(* IEC 61131-3 sources: plcfuzz/testcases/beremiz_projects/random_projects (part 4) *)

(* Additional processing to handle clocks - in CODESYS, it only starts
    with rising edge and can not be placed inside IF statement *)
IF(t0_up = TRUE) THEN
    t0_reset := TRUE;
ELSIF(t0_start = TRUE AND t0_up = FALSE) THEN
    t0_up := TRUE;  t0_reset := FALSE;
END_IF
t0(IN:=t0_reset, PT:=T0_VALUE);

END_FUNCTION_BLOCK

(* ---- IndustrialAuto2.st ---- *)
FUNCTION_BLOCK FB_G4LTL

   (* Variable definition *)
   VAR_INPUT
      x0	: BOOL;
      x1	: BOOL;
   END_VAR
   VAR_OUTPUT
      y0	: BOOL;
   END_VAR
   VAR
   (* The total number of states equals to 1 *)
      cstate6	: LINT := 0;
   END_VAR

   (* Control logic *)
CASE cstate6 OF
0:
    IF ((x0 = FALSE) AND  (x1 = TRUE)) OR ((x0 = TRUE) AND  (x1 = FALSE)) THEN
        cstate6 := 0; y0 := FALSE;
    ELSIF ((x0 = FALSE) AND  (x1 = FALSE)) OR ((x0 = TRUE) AND  (x1 = TRUE)) THEN
        cstate6 := 0; y0 := TRUE;
    END_IF;
END_CASE;

END_FUNCTION_BLOCK

(* ---- IndustrialAuto3.st ---- *)
FUNCTION_BLOCK FB_G4LTL

   (* Variable definition *)
   VAR_INPUT
      x0	: BOOL;
      x1	: BOOL;
      x2	: BOOL;
      x3	: BOOL;
   END_VAR
   VAR_OUTPUT
      y0	: BOOL;
   END_VAR
   VAR
   (* The total number of states equals to 12 *)
      cstate3	: LINT := 0;
   END_VAR

   (* Control logic *)
CASE cstate3 OF
22:
    IF ((x0 = TRUE) AND  (x1 = TRUE) AND  (x2 = TRUE) AND  (x3 = FALSE)) THEN
        cstate3 := 247; y0 := FALSE;
    ELSIF ((x0 = FALSE) AND  ( TRUE ) AND  ( TRUE ) AND  ( TRUE )) OR ((x0 = TRUE) AND  ( TRUE ) AND  (x2 = FALSE) AND  ( TRUE )) THEN
        cstate3 := 22; y0 := FALSE;
    ELSIF ((x0 = TRUE) AND  (x1 = FALSE) AND  (x2 = TRUE) AND  (x3 = FALSE)) THEN
        cstate3 := 246; y0 := TRUE;
    ELSIF ((x0 = TRUE) AND  ( TRUE ) AND  (x2 = TRUE) AND  (x3 = TRUE)) THEN
        cstate3 := 29; y0 := FALSE;
    END_IF;
0:
    IF ((x0 = FALSE) AND  (x1 = FALSE) AND  (x2 = TRUE) AND  (x3 = FALSE)) THEN
        cstate3 := 0; y0 := FALSE;
    ELSIF ((x0 = FALSE) AND  (x1 = TRUE) AND  (x2 = TRUE) AND  (x3 = FALSE)) THEN
        cstate3 := 24; y0 := FALSE;
    ELSIF ((x0 = FALSE) AND  (x1 = TRUE) AND  ( TRUE ) AND  (x3 = TRUE)) OR ((x0 = TRUE) AND  (x1 = TRUE) AND  (x2 = FALSE) AND  (x3 = TRUE)) THEN
        cstate3 := 22; y0 := FALSE;
    ELSIF ((x0 = TRUE) AND  (x1 = TRUE) AND  (x2 = TRUE) AND  (x3 = FALSE)) THEN
        cstate3 := 28; y0 := FALSE;
    ELSIF (( TRUE ) AND  (x1 = TRUE) AND  (x2 = FALSE) AND  (x3 = FALSE)) THEN
        cstate3 := 20; y0 := FALSE;
    ELSIF ((x0 = TRUE) AND  (x1 = FALSE) AND  (x2 = TRUE) AND  (x3 = FALSE)) THEN
        cstate3 := 27; y0 := TRUE;
    ELSIF ((x0 = TRUE) AND  (x1 = TRUE) AND  (x2 = TRUE) AND  (x3 = TRUE)) THEN
        cstate3 := 29; y0 := FALSE;
    ELSIF (( TRUE ) AND  (x1 = FALSE) AND  (x2 = FALSE) AND  ( TRUE )) OR (( TRUE ) AND  (x1 = FALSE) AND  (x2 = TRUE) AND  (x3 = TRUE)) THEN
        cstate3 := 18; y0 := FALSE;
    END_IF;
243:
    IF ((x0 = FALSE) AND  (x1 = FALSE) AND  (x2 = TRUE) AND  (x3 = TRUE)) OR ((x0 = TRUE) AND  ( TRUE ) AND  (x2 = TRUE) AND  (x3 = TRUE)) THEN
        cstate3 := 29; y0 := FALSE;
    ELSIF (( TRUE ) AND  ( TRUE ) AND  (x2 = FALSE) AND  (x3 = FALSE)) THEN
        cstate3 := 20; y0 := FALSE;
    ELSIF ((x0 = FALSE) AND  (x1 = FALSE) AND  (x2 = FALSE) AND  (x3 = TRUE)) OR ((x0 = FALSE) AND  (x1 = TRUE) AND  ( TRUE ) AND  (x3 = TRUE)) OR ((x0 = TRUE) AND  ( TRUE ) AND  (x2 = FALSE) AND  (x3 = TRUE)) THEN
        cstate3 := 22; y0 := FALSE;
    ELSIF ((x0 = FALSE) AND  (x1 = TRUE) AND  (x2 = TRUE) AND  (x3 = FALSE)) THEN
        cstate3 := 24; y0 := FALSE;
    ELSIF ((x0 = TRUE) AND  (x1 = TRUE) AND  (x2 = TRUE) AND  (x3 = FALSE)) THEN
        cstate3 := 28; y0 := FALSE;
    ELSIF (( TRUE ) AND  (x1 = FALSE) AND  (x2 = TRUE) AND  (x3 = FALSE)) THEN
        cstate3 := 243; y0 := TRUE;
    END_IF;
24:
    IF ((x0 = TRUE) AND  ( TRUE ) AND  (x2 = TRUE) AND  (x3 = TRUE)) THEN
        cstate3 := 29; y0 := FALSE;
    ELSIF (( TRUE ) AND  ( TRUE ) AND  (x2 = FALSE) AND  (x3 = FALSE)) THEN
        cstate3 := 20; y0 := FALSE;
    ELSIF ((x0 = FALSE) AND  ( TRUE ) AND  ( TRUE ) AND  (x3 = TRUE)) OR ((x0 = TRUE) AND  ( TRUE ) AND  (x2 = FALSE) AND  (x3 = TRUE)) THEN
        cstate3 := 22; y0 := FALSE;
    ELSIF ((x0 = TRUE) AND  (x1 = TRUE) AND  (x2 = TRUE) AND  (x3 = FALSE)) THEN
        cstate3 := 28; y0 := FALSE;
    ELSIF ((x0 = TRUE) AND  (x1 = FALSE) AND  (x2 = TRUE) AND  (x3 = FALSE)) THEN
        cstate3 := 243; y0 := TRUE;
    ELSIF ((x0 = FALSE) AND  ( TRUE ) AND  (x2 = TRUE) AND  (x3 = FALSE)) THEN
        cstate3 := 24; y0 := FALSE;
    END_IF;
246:
    IF ((x0 = FALSE) AND  (x1 = FALSE) AND  (x2 = FALSE) AND  ( TRUE )) OR ((x0 = FALSE) AND  (x1 = TRUE) AND  (x2 = FALSE) AND  ( TRUE )) OR ((x0 = FALSE) AND  (x1 = TRUE) AND  (x2 = TRUE) AND  (x3 = TRUE)) OR ((x0 = TRUE) AND  ( TRUE ) AND  (x2 = FALSE) AND  ( TRUE )) THEN
        cstate3 := 22; y0 := FALSE;
    ELSIF (( TRUE ) AND  (x1 = FALSE) AND  (x2 = TRUE) AND  (x3 = FALSE)) THEN
        cstate3 := 246; y0 := TRUE;
    ELSIF ((x0 = FALSE) AND  (x1 = FALSE) AND  (x2 = TRUE) AND  (x3 = TRUE)) OR ((x0 = TRUE) AND  ( TRUE ) AND  (x2 = TRUE) AND  (x3 = TRUE)) THEN
        cstate3 := 29; y0 := FALSE;
    ELSIF ((x0 = FALSE) AND  (x1 = TRUE) AND  (x2 = TRUE) AND  (x3 = FALSE)) THEN
        cstate3 := 786; y0 := FALSE;
    ELSIF ((x0 = TRUE) AND  (x1 = TRUE) AND  (x2 = TRUE) AND  (x3 = FALSE)) THEN
        cstate3 := 247; y0 := FALSE;
    END_IF;
27:
    IF ((x0 = FALSE) AND  (x1 = TRUE) AND  (x2 = TRUE) AND  (x3 = FALSE)) THEN
        cstate3 := 24; y0 := FALSE;
    ELSIF (( TRUE ) AND  (x1 = TRUE) AND  (x2 = FALSE) AND  (x3 = FALSE)) THEN
        cstate3 := 20; y0 := FALSE;
    ELSIF ((x0 = FALSE) AND  (x1 = TRUE) AND  ( TRUE ) AND  (x3 = TRUE)) OR ((x0 = TRUE) AND  (x1 = TRUE) AND  (x2 = FALSE) AND  (x3 = TRUE)) THEN
        cstate3 := 22; y0 := FALSE;
    ELSIF ((x0 = TRUE) AND  (x1 = TRUE) AND  (x2 = TRUE) AND  (x3 = FALSE)) THEN
        cstate3 := 28; y0 := FALSE;
    ELSIF (( TRUE ) AND  (x1 = FALSE) AND  (x2 = TRUE) AND  (x3 = FALSE)) THEN
        cstate3 := 27; y0 := TRUE;
    ELSIF ((x0 = TRUE) AND  (x1 = TRUE) AND  (x2 = TRUE) AND  (x3 = TRUE)) THEN
        cstate3 := 29; y0 := FALSE;
    ELSIF (( TRUE ) AND  (x1 = FALSE) AND  (x2 = FALSE) AND  ( TRUE )) OR (( TRUE ) AND  (x1 = FALSE) AND  (x2 = TRUE) AND  (x3 = TRUE)) THEN
        cstate3 := 18; y0 := FALSE;
    END_IF;
247:
    IF ((x0 = FALSE) AND  (x1 = TRUE) AND  (x2 = TRUE) AND  (x3 = FALSE)) THEN
        cstate3 := 786; y0 := FALSE;
    ELSIF ((x0 = FALSE) AND  (x1 = FALSE) AND  (x2 = TRUE) AND  (x3 = FALSE)) OR ((x0 = TRUE) AND  (x1 = TRUE) AND  (x2 = TRUE) AND  (x3 = FALSE)) THEN
        cstate3 := 247; y0 := FALSE;
    ELSIF ((x0 = FALSE) AND  (x1 = FALSE) AND  (x2 = FALSE) AND  ( TRUE )) OR ((x0 = FALSE) AND  (x1 = TRUE) AND  (x2 = FALSE) AND  ( TRUE )) OR ((x0 = FALSE) AND  (x1 = TRUE) AND  (x2 = TRUE) AND  (x3 = TRUE)) OR ((x0 = TRUE) AND  ( TRUE ) AND  (x2 = FALSE) AND  ( TRUE )) THEN
        cstate3 := 22; y0 := FALSE;
    ELSIF ((x0 = TRUE) AND  (x1 = FALSE) AND  (x2 = TRUE) AND  (x3 = FALSE)) THEN
        cstate3 := 246; y0 := TRUE;
    ELSIF ((x0 = FALSE) AND  (x1 = FALSE) AND  (x2 = TRUE) AND  (x3 = TRUE)) OR ((x0 = TRUE) AND  ( TRUE ) AND  (x2 = TRUE) AND  (x3 = TRUE)) THEN
        cstate3 := 29; y0 := FALSE;
    END_IF;
786:
    IF ((x0 = TRUE) AND  (x1 = TRUE) AND  (x2 = TRUE) AND  (x3 = FALSE)) THEN
        cstate3 := 247; y0 := FALSE;
    ELSIF ((x0 = FALSE) AND  ( TRUE ) AND  (x2 = FALSE) AND  ( TRUE )) OR ((x0 = FALSE) AND  ( TRUE ) AND  (x2 = TRUE) AND  (x3 = TRUE)) OR ((x0 = TRUE) AND  ( TRUE ) AND  (x2 = FALSE) AND  ( TRUE )) THEN
        cstate3 := 22; y0 := FALSE;
    ELSIF ((x0 = FALSE) AND  ( TRUE ) AND  (x2 = TRUE) AND  (x3 = FALSE)) THEN
        cstate3 := 786; y0 := FALSE;
    ELSIF ((x0 = TRUE) AND  (x1 = FALSE) AND  (x2 = TRUE) AND  (x3 = FALSE)) THEN
        cstate3 := 246; y0 := TRUE;
    ELSIF ((x0 = TRUE) AND  ( TRUE ) AND  (x2 = TRUE) AND  (x3 = TRUE)) THEN
        cstate3 := 29; y0 := FALSE;
    END_IF;
28:
    IF ((x0 = FALSE) AND  (x1 = FALSE) AND  (x2 = TRUE) AND  (x3 = FALSE)) OR ((x0 = TRUE) AND  (x1 = TRUE) AND  (x2 = TRUE) AND  (x3 = FALSE)) THEN
        cstate3 := 28; y0 := FALSE;
    ELSIF (( TRUE ) AND  ( TRUE ) AND  (x2 = FALSE) AND  (x3 = FALSE)) THEN
        cstate3 := 20; y0 := FALSE;
    ELSIF ((x0 = FALSE) AND  (x1 = FALSE) AND  (x2 = FALSE) AND  (x3 = TRUE)) OR ((x0 = FALSE) AND  (x1 = TRUE) AND  ( TRUE ) AND  (x3 = TRUE)) OR ((x0 = TRUE) AND  ( TRUE ) AND  (x2 = FALSE) AND  (x3 = TRUE)) THEN
        cstate3 := 22; y0 := FALSE;
    ELSIF ((x0 = FALSE) AND  (x1 = TRUE) AND  (x2 = TRUE) AND  (x3 = FALSE)) THEN
        cstate3 := 24; y0 := FALSE;
    ELSIF ((x0 = TRUE) AND  (x1 = FALSE) AND  (x2 = TRUE) AND  (x3 = FALSE)) THEN
        cstate3 := 243; y0 := TRUE;
    ELSIF ((x0 = FALSE) AND  (x1 = FALSE) AND  (x2 = TRUE) AND  (x3 = TRUE)) OR ((x0 = TRUE) AND  ( TRUE ) AND  (x2 = TRUE) AND  (x3 = TRUE)) THEN
        cstate3 := 29; y0 := FALSE;
    END_IF;
29:
    IF ((x0 = TRUE) AND  (x1 = TRUE) AND  (x2 = TRUE) AND  (x3 = FALSE)) THEN
        cstate3 := 247; y0 := FALSE;
    ELSIF ((x0 = FALSE) AND  (x1 = FALSE) AND  (x2 = TRUE) AND  ( TRUE )) OR ((x0 = TRUE) AND  ( TRUE ) AND  (x2 = TRUE) AND  (x3 = TRUE)) THEN
        cstate3 := 29; y0 := FALSE;
    ELSIF ((x0 = TRUE) AND  (x1 = FALSE) AND  (x2 = TRUE) AND  (x3 = FALSE)) THEN
        cstate3 := 246; y0 := TRUE;
    ELSIF ((x0 = FALSE) AND  (x1 = FALSE) AND  (x2 = FALSE) AND  ( TRUE )) OR ((x0 = FALSE) AND  (x1 = TRUE) AND  ( TRUE ) AND  ( TRUE )) OR ((x0 = TRUE) AND  ( TRUE ) AND  (x2 = FALSE) AND  ( TRUE )) THEN
        cstate3 := 22; y0 := FALSE;
    END_IF;
18:
    IF ((x0 = TRUE) AND  (x1 = TRUE) AND  (x2 = TRUE) AND  (x3 = TRUE)) THEN
        cstate3 := 29; y0 := FALSE;
    ELSIF ((x0 = TRUE) AND  (x1 = FALSE) AND  (x2 = TRUE) AND  (x3 = FALSE)) THEN
        cstate3 := 27; y0 := TRUE;
    ELSIF ((x0 = FALSE) AND  (x1 = FALSE) AND  ( TRUE ) AND  ( TRUE )) OR ((x0 = TRUE) AND  (x1 = FALSE) AND  (x2 = FALSE) AND  ( TRUE )) OR ((x0 = TRUE) AND  (x1 = FALSE) AND  (x2 = TRUE) AND  (x3 = TRUE)) THEN
        cstate3 := 18; y0 := FALSE;
    ELSIF ((x0 = FALSE) AND  (x1 = TRUE) AND  ( TRUE ) AND  (x3 = FALSE)) OR ((x0 = TRUE) AND  (x1 = TRUE) AND  (x2 = FALSE) AND  (x3 = FALSE)) THEN
        cstate3 := 20; y0 := FALSE;
    ELSIF ((x0 = FALSE) AND  (x1 = TRUE) AND  ( TRUE ) AND  (x3 = TRUE)) OR ((x0 = TRUE) AND  (x1 = TRUE) AND  (x2 = FALSE) AND  (x3 = TRUE)) THEN
        cstate3 := 22; y0 := FALSE;
    ELSIF ((x0 = TRUE) AND  (x1 = TRUE) AND  (x2 = TRUE) AND  (x3 = FALSE)) THEN
        cstate3 := 28; y0 := FALSE;
    END_IF;
20:
    IF ((x0 = TRUE) AND  ( TRUE ) AND  (x2 = TRUE) AND  (x3 = TRUE)) THEN
        cstate3 := 29; y0 := FALSE;
    ELSIF ((x0 = FALSE) AND  ( TRUE ) AND  ( TRUE ) AND  (x3 = TRUE)) OR ((x0 = TRUE) AND  ( TRUE ) AND  (x2 = FALSE) AND  (x3 = TRUE)) THEN
        cstate3 := 22; y0 := FALSE;
    ELSIF ((x0 = FALSE) AND  ( TRUE ) AND  ( TRUE ) AND  (x3 = FALSE)) OR ((x0 = TRUE) AND  ( TRUE ) AND  (x2 = FALSE) AND  (x3 = FALSE)) THEN
        cstate3 := 20; y0 := FALSE;
    ELSIF ((x0 = TRUE) AND  (x1 = TRUE) AND  (x2 = TRUE) AND  (x3 = FALSE)) THEN
        cstate3 := 28; y0 := FALSE;
    ELSIF ((x0 = TRUE) AND  (x1 = FALSE) AND  (x2 = TRUE) AND  (x3 = FALSE)) THEN
        cstate3 := 243; y0 := TRUE;
    END_IF;
END_CASE;

END_FUNCTION_BLOCK

(* ---- IndustrialAuto4.st ---- *)
FUNCTION_BLOCK FB_G4LTL

   (* Variable definition *)
   VAR_INPUT
      x0	: BOOL;
      x1	: BOOL;
      x2	: BOOL;
      x3	: BOOL;
   END_VAR
   VAR_OUTPUT
      y0	: BOOL;
      y1	: BOOL;
   END_VAR
   VAR
   (* The total number of states equals to 2 *)
      cstate21	: LINT := 0;
   END_VAR

   (* Control logic *)
CASE cstate21 OF
0:
    IF ((x0 = FALSE) AND  (x1 = FALSE) AND  (x2 = FALSE) AND  (x3 = TRUE)) THEN
        cstate21 := 0; y0 := FALSE; y1 := FALSE;
    ELSIF ((x0 = FALSE) AND  (x1 = TRUE) AND  ( TRUE ) AND  (x3 = TRUE)) OR ((x0 = TRUE) AND  (x1 = FALSE) AND  (x2 = TRUE) AND  ( TRUE )) OR ((x0 = TRUE) AND  (x1 = TRUE) AND  (x2 = FALSE) AND  (x3 = TRUE)) OR ((x0 = TRUE) AND  (x1 = TRUE) AND  (x2 = TRUE) AND  ( TRUE )) THEN
        cstate21 := 1; y0 := FALSE; y1 := FALSE;
    ELSIF ((x0 = FALSE) AND  (x1 = FALSE) AND  (x2 = FALSE) AND  (x3 = FALSE)) OR ((x0 = FALSE) AND  (x1 = FALSE) AND  (x2 = TRUE) AND  ( TRUE )) OR ((x0 = FALSE) AND  (x1 = TRUE) AND  ( TRUE ) AND  (x3 = FALSE)) THEN
        cstate21 := 0; y0 := FALSE; y1 := FALSE;
    ELSIF ((x0 = TRUE) AND  (x1 = TRUE) AND  (x2 = FALSE) AND  (x3 = FALSE)) THEN
        cstate21 := 0; y0 := TRUE; y1 := TRUE;
    ELSIF ((x0 = TRUE) AND  (x1 = FALSE) AND  (x2 = FALSE) AND  (x3 = TRUE)) THEN
        cstate21 := 0; y0 := TRUE; y1 := FALSE;
    ELSIF ((x0 = TRUE) AND  (x1 = FALSE) AND  (x2 = FALSE) AND  (x3 = FALSE)) THEN
        cstate21 := 0; y0 := TRUE; y1 := FALSE;
    END_IF;
1:
    IF ((x0 = TRUE) AND  (x1 = FALSE) AND  (x2 = FALSE) AND  ( TRUE )) OR ((x0 = TRUE) AND  (x1 = TRUE) AND  (x2 = FALSE) AND  (x3 = FALSE)) THEN
        cstate21 := 1; y0 := FALSE; y1 := FALSE;
    ELSIF ((x0 = FALSE) AND  (x1 = FALSE) AND  (x2 = FALSE) AND  (x3 = FALSE)) OR ((x0 = FALSE) AND  (x1 = FALSE) AND  (x2 = TRUE) AND  ( TRUE )) OR ((x0 = FALSE) AND  (x1 = TRUE) AND  ( TRUE ) AND  (x3 = FALSE)) THEN
        cstate21 := 1; y0 := FALSE; y1 := FALSE;
    ELSIF ((x0 = FALSE) AND  (x1 = TRUE) AND  ( TRUE ) AND  (x3 = TRUE)) OR ((x0 = TRUE) AND  (x1 = FALSE) AND  (x2 = TRUE) AND  ( TRUE )) OR ((x0 = TRUE) AND  (x1 = TRUE) AND  (x2 = FALSE) AND  (x3 = TRUE)) OR ((x0 = TRUE) AND  (x1 = TRUE) AND  (x2 = TRUE) AND  ( TRUE )) THEN
        cstate21 := 1; y0 := FALSE; y1 := FALSE;
    ELSIF ((x0 = FALSE) AND  (x1 = FALSE) AND  (x2 = FALSE) AND  (x3 = TRUE)) THEN
        cstate21 := 1; y0 := FALSE; y1 := FALSE;
    END_IF;
END_CASE;

END_FUNCTION_BLOCK

(* ---- IndustrialAuto5.st ---- *)
FUNCTION_BLOCK FB_G4LTL

   (* Variable definition *)
   VAR_INPUT
      x0	: BOOL;
      x1	: BOOL;
      c1_geq500	: BOOL;
   END_VAR
   VAR_OUTPUT
      y0	: BOOL;
      c1_add1	: BOOL;
      c1_reset	: BOOL;
   END_VAR
   VAR
   (* The total number of states equals to 4 *)
      cstate18	: LINT := 0;
   END_VAR

   (* Control logic *)
CASE cstate18 OF
0:
    IF ((x0 = FALSE) AND  (x1 = TRUE) AND  (c1_geq500 = TRUE)) THEN
        cstate18 := 3; y0 := TRUE; c1_add1 := FALSE; c1_reset := TRUE;
    ELSIF ((x0 = FALSE) AND  (x1 = FALSE) AND  (c1_geq500 = TRUE)) THEN
        cstate18 := 3; y0 := TRUE; c1_add1 := FALSE; c1_reset := FALSE;
    ELSIF ((x0 = FALSE) AND  (x1 = TRUE) AND  (c1_geq500 = FALSE)) THEN
        cstate18 := 3; y0 := FALSE; c1_add1 := FALSE; c1_reset := TRUE;
    ELSIF ((x0 = FALSE) AND  (x1 = FALSE) AND  (c1_geq500 = FALSE)) THEN
        cstate18 := 3; y0 := FALSE; c1_add1 := FALSE; c1_reset := FALSE;
    ELSIF ((x0 = TRUE) AND  (x1 = TRUE) AND  ( TRUE )) THEN
        cstate18 := 1; y0 := FALSE; c1_add1 := FALSE; c1_reset := FALSE;
    ELSIF ((x0 = TRUE) AND  (x1 = FALSE) AND  (c1_geq500 = TRUE)) THEN
        cstate18 := 2; y0 := TRUE; c1_add1 := TRUE; c1_reset := FALSE;
    ELSIF ((x0 = TRUE) AND  (x1 = FALSE) AND  (c1_geq500 = FALSE)) THEN
        cstate18 := 2; y0 := FALSE; c1_add1 := TRUE; c1_reset := FALSE;
    END_IF;
1:
    IF ((x0 = TRUE) AND  (x1 = TRUE) AND  ( TRUE )) THEN
        cstate18 := 1; y0 := FALSE; c1_add1 := FALSE; c1_reset := FALSE;
    ELSIF ((x0 = FALSE) AND  ( TRUE ) AND  (c1_geq500 = FALSE)) OR ((x0 = TRUE) AND  (x1 = FALSE) AND  (c1_geq500 = FALSE)) THEN
        cstate18 := 1; y0 := FALSE; c1_add1 := FALSE; c1_reset := FALSE;
    ELSIF ((x0 = FALSE) AND  ( TRUE ) AND  (c1_geq500 = TRUE)) OR ((x0 = TRUE) AND  (x1 = FALSE) AND  (c1_geq500 = TRUE)) THEN
        cstate18 := 1; y0 := FALSE; c1_add1 := FALSE; c1_reset := FALSE;
    END_IF;
2:
    IF ((x0 = TRUE) AND  (x1 = TRUE) AND  ( TRUE )) THEN
        cstate18 := 1; y0 := FALSE; c1_add1 := FALSE; c1_reset := FALSE;
    ELSIF ((x0 = FALSE) AND  (x1 = FALSE) AND  (c1_geq500 = TRUE)) THEN
        cstate18 := 3; y0 := TRUE; c1_add1 := FALSE; c1_reset := FALSE;
    ELSIF ((x0 = FALSE) AND  (x1 = TRUE) AND  (c1_geq500 = FALSE)) THEN
        cstate18 := 3; y0 := FALSE; c1_add1 := FALSE; c1_reset := TRUE;
    ELSIF ((x0 = FALSE) AND  (x1 = TRUE) AND  (c1_geq500 = TRUE)) THEN
        cstate18 := 3; y0 := TRUE; c1_add1 := FALSE; c1_reset := TRUE;
    ELSIF ((x0 = FALSE) AND  (x1 = FALSE) AND  (c1_geq500 = FALSE)) THEN
        cstate18 := 3; y0 := FALSE; c1_add1 := FALSE; c1_reset := FALSE;
    ELSIF ((x0 = TRUE) AND  (x1 = FALSE) AND  (c1_geq500 = FALSE)) THEN
        cstate18 := 2; y0 := FALSE; c1_add1 := FALSE; c1_reset := FALSE;
    ELSIF ((x0 = TRUE) AND  (x1 = FALSE) AND  (c1_geq500 = TRUE)) THEN
        cstate18 := 2; y0 := TRUE; c1_add1 := FALSE; c1_reset := FALSE;
    END_IF;
3:
    IF ((x0 = FALSE) AND  (x1 = FALSE) AND  (c1_geq500 = FALSE)) THEN
        cstate18 := 3; y0 := FALSE; c1_add1 := FALSE; c1_reset := FALSE;
    ELSIF ((x0 = FALSE) AND  (x1 = FALSE) AND  (c1_geq500 = TRUE)) THEN
        cstate18 := 3; y0 := TRUE; c1_add1 := FALSE; c1_reset := FALSE;
    ELSIF ((x0 = FALSE) AND  (x1 = TRUE) AND  (c1_geq500 = FALSE)) THEN
        cstate18 := 3; y0 := FALSE; c1_add1 := FALSE; c1_reset := TRUE;
    ELSIF ((x0 = FALSE) AND  (x1 = TRUE) AND  (c1_geq500 = TRUE)) THEN
        cstate18 := 3; y0 := TRUE; c1_add1 := FALSE; c1_reset := TRUE;
    ELSIF ((x0 = TRUE) AND  (x1 = TRUE) AND  ( TRUE )) THEN
        cstate18 := 1; y0 := FALSE; c1_add1 := FALSE; c1_reset := FALSE;
    ELSIF ((x0 = TRUE) AND  (x1 = FALSE) AND  (c1_geq500 = FALSE)) THEN
        cstate18 := 2; y0 := FALSE; c1_add1 := TRUE; c1_reset := FALSE;
    ELSIF ((x0 = TRUE) AND  (x1 = FALSE) AND  (c1_geq500 = TRUE)) THEN
        cstate18 := 2; y0 := TRUE; c1_add1 := TRUE; c1_reset := FALSE;
    END_IF;
END_CASE;

END_FUNCTION_BLOCK

(* ---- IndustrialAuto6.st ---- *)
FUNCTION_BLOCK FB_G4LTL

   (* Variable definition *)
   VAR_INPUT
      x1	: BOOL;
   END_VAR
   VAR_OUTPUT
      y1	: BOOL;
   END_VAR
   VAR
   (* The total number of states equals to 7 *)
      cstate12	: LINT := 0;
      t	: TON;
      t_reset	: BOOL := FALSE;
      t_up	: BOOL := FALSE;
      t_start	: BOOL := FALSE;
   END_VAR

   (* Constant definition (depending on compiler, one might need to move to normal variables) *)

   (* Each time constant has a difference of 1 period (cycle-time); please substract it when needed  *)
   VAR CONST
      T_VALUE	: TIME := TIME#5s;
   END_VAR

   (* Control logic *)
CASE cstate12 OF
0:
    IF ((x1 = FALSE) AND  (t.Q = FALSE)) THEN
        cstate12 := 1; y1 := FALSE; t_start := FALSE;
    ELSIF ((x1 = TRUE) AND  ( TRUE )) THEN
        cstate12 := 3; y1 := TRUE; t_start := FALSE;
    ELSIF ((x1 = FALSE) AND  (t.Q = TRUE)) THEN
        cstate12 := 5; y1 := FALSE; t_start := FALSE;
    END_IF;
1:
    IF ((x1 = FALSE) AND  (t.Q = FALSE)) THEN
        cstate12 := 1; y1 := FALSE; t_start := FALSE;
    ELSIF ((x1 = FALSE) AND  (t.Q = TRUE)) THEN
        cstate12 := 5; y1 := FALSE; t_start := FALSE;
    ELSIF ((x1 = TRUE) AND  ( TRUE )) THEN
        cstate12 := 3; y1 := TRUE; t_start := FALSE;
    END_IF;
2:
    IF ((x1 = TRUE) AND  (t.Q = FALSE)) THEN
        cstate12 := 2; y1 := TRUE; t_start := FALSE;
    ELSIF ((x1 = TRUE) AND  (t.Q = TRUE)) THEN
        cstate12 := 3; y1 := TRUE; t_start := FALSE;
    ELSIF ((x1 = FALSE) AND  (t.Q = FALSE)) THEN
        cstate12 := 4; y1 := TRUE; t_start := TRUE; t_up := FALSE;
    ELSIF ((x1 = FALSE) AND  (t.Q = TRUE)) THEN
        cstate12 := 6; y1 := TRUE; t_start := TRUE; t_up := FALSE;
    END_IF;
3:
    IF ((x1 = FALSE) AND  (t.Q = TRUE)) THEN
        cstate12 := 6; y1 := TRUE; t_start := TRUE; t_up := FALSE;
    ELSIF ((x1 = FALSE) AND  (t.Q = FALSE)) THEN
        cstate12 := 4; y1 := TRUE; t_start := TRUE; t_up := FALSE;
    ELSIF ((x1 = TRUE) AND  ( TRUE )) THEN
        cstate12 := 3; y1 := TRUE; t_start := FALSE;
    END_IF;
4:
    IF ((x1 = FALSE) AND  (t.Q = TRUE)) THEN
        cstate12 := 5; y1 := FALSE; t_start := FALSE;
    ELSIF ((x1 = FALSE) AND  (t.Q = FALSE)) THEN
        cstate12 := 4; y1 := TRUE; t_start := FALSE;
    ELSIF ((x1 = TRUE) AND  (t.Q = FALSE)) THEN
        cstate12 := 2; y1 := TRUE; t_start := FALSE;
    ELSIF ((x1 = TRUE) AND  (t.Q = TRUE)) THEN
        cstate12 := 3; y1 := TRUE; t_start := FALSE;
    END_IF;
5:
    IF ((x1 = TRUE) AND  ( TRUE )) THEN
        cstate12 := 3; y1 := TRUE; t_start := FALSE;
    ELSIF ((x1 = FALSE) AND  (t.Q = FALSE)) THEN
        cstate12 := 1; y1 := FALSE; t_start := FALSE;
    ELSIF ((x1 = FALSE) AND  (t.Q = TRUE)) THEN
        cstate12 := 5; y1 := FALSE; t_start := FALSE;
    END_IF;
6:
    IF ((x1 = FALSE) AND  (t.Q = TRUE)) THEN
        cstate12 := 5; y1 := FALSE; t_start := FALSE;
    ELSIF ((x1 = FALSE) AND  (t.Q = FALSE)) THEN
        cstate12 := 4; y1 := TRUE; t_start := FALSE;
    ELSIF ((x1 = TRUE) AND  (t.Q = FALSE)) THEN
        cstate12 := 2; y1 := TRUE; t_start := FALSE;
    ELSIF ((x1 = TRUE) AND  (t.Q = TRUE)) THEN
        cstate12 := 3; y1 := TRUE; t_start := FALSE;
    END_IF;
END_CASE;

(* Additional processing to handle clocks - in CODESYS, it only starts
    with rising edge and can not be placed inside IF statement *)
IF(t_up = TRUE) THEN
    t_reset := TRUE;
ELSIF(t_start = TRUE AND t_up = FALSE) THEN
    t_up := TRUE;  t_reset := FALSE;
END_IF
t(IN:=t_reset, PT:=T_VALUE);

END_FUNCTION_BLOCK

(* ---- IndustrialAuto7.st ---- *)
FUNCTION_BLOCK FB_G4LTL

   (* Variable definition *)
   VAR_INPUT
      x1	: BOOL;
   END_VAR
   VAR_OUTPUT
      y1	: BOOL;
   END_VAR
   VAR
   (* The total number of states equals to 7 *)
      cstate71	: LINT := 0;
      t	: TON;
      t_reset	: BOOL := FALSE;
      t_up	: BOOL := FALSE;
      t_start	: BOOL := FALSE;
   END_VAR

   (* Constant definition (depending on compiler, one might need to move to normal variables) *)

   (* Each time constant has a difference of 1 period (cycle-time); please substract it when needed  *)
   VAR CONST
      T_VALUE	: TIME := TIME#3s;
   END_VAR

   (* Control logic *)
CASE cstate71 OF
0:
    IF ((x1 = TRUE) AND  (t.Q = FALSE)) THEN
        cstate71 := 2; y1 := FALSE; t_start := FALSE;
    ELSIF ((x1 = FALSE) AND  ( TRUE )) THEN
        cstate71 := 6; y1 := FALSE; t_start := FALSE;
    ELSIF ((x1 = TRUE) AND  (t.Q = TRUE)) THEN
        cstate71 := 2; y1 := TRUE; t_start := FALSE;
    END_IF;
1:
    IF ((x1 = TRUE) AND  (t.Q = TRUE)) THEN
        cstate71 := 2; y1 := TRUE; t_start := FALSE;
    ELSIF ((x1 = TRUE) AND  (t.Q = FALSE)) THEN
        cstate71 := 1; y1 := FALSE; t_start := FALSE;
    ELSIF ((x1 = FALSE) AND  (t.Q = TRUE)) THEN
        cstate71 := 6; y1 := FALSE; t_start := FALSE;
    ELSIF ((x1 = FALSE) AND  (t.Q = FALSE)) THEN
        cstate71 := 5; y1 := FALSE; t_start := FALSE;
    END_IF;
2:
    IF ((x1 = TRUE) AND  (t.Q = FALSE)) THEN
        cstate71 := 2; y1 := FALSE; t_start := FALSE;
    ELSIF ((x1 = TRUE) AND  (t.Q = TRUE)) THEN
        cstate71 := 2; y1 := TRUE; t_start := FALSE;
    ELSIF ((x1 = FALSE) AND  ( TRUE )) THEN
        cstate71 := 6; y1 := FALSE; t_start := FALSE;
    END_IF;
3:
    IF ((x1 = TRUE) AND  (t.Q = FALSE)) THEN
        cstate71 := 3; y1 := FALSE; t_start := FALSE;
    ELSIF ((x1 = FALSE) AND  (t.Q = FALSE)) THEN
        cstate71 := 4; y1 := FALSE; t_start := FALSE;
    ELSIF ((x1 = TRUE) AND  (t.Q = TRUE)) THEN
        cstate71 := 2; y1 := TRUE; t_start := FALSE;
    ELSIF ((x1 = FALSE) AND  (t.Q = TRUE)) THEN
        cstate71 := 6; y1 := FALSE; t_start := FALSE;
    END_IF;
4:
    IF ((x1 = FALSE) AND  (t.Q = FALSE)) THEN
        cstate71 := 4; y1 := FALSE; t_start := FALSE;
    ELSIF ((x1 = FALSE) AND  (t.Q = TRUE)) THEN
        cstate71 := 6; y1 := FALSE; t_start := FALSE;
    ELSIF ((x1 = TRUE) AND  (t.Q = FALSE)) THEN
        cstate71 := 3; y1 := FALSE; t_start := TRUE; t_up := FALSE;
    ELSIF ((x1 = TRUE) AND  (t.Q = TRUE)) THEN
        cstate71 := 1; y1 := TRUE; t_start := TRUE; t_up := FALSE;
    END_IF;
5:
    IF ((x1 = FALSE) AND  (t.Q = TRUE)) THEN
        cstate71 := 6; y1 := FALSE; t_start := FALSE;
    ELSIF ((x1 = FALSE) AND  (t.Q = FALSE)) THEN
        cstate71 := 5; y1 := FALSE; t_start := FALSE;
    ELSIF ((x1 = TRUE) AND  (t.Q = TRUE)) THEN
        cstate71 := 1; y1 := TRUE; t_start := TRUE; t_up := FALSE;
    ELSIF ((x1 = TRUE) AND  (t.Q = FALSE)) THEN
        cstate71 := 3; y1 := FALSE; t_start := TRUE; t_up := FALSE;
    END_IF;
6:
    IF ((x1 = TRUE) AND  (t.Q = TRUE)) THEN
        cstate71 := 1; y1 := TRUE; t_start := TRUE; t_up := FALSE;
    ELSIF ((x1 = TRUE) AND  (t.Q = FALSE)) THEN
        cstate71 := 3; y1 := FALSE; t_start := TRUE; t_up := FALSE;
    ELSIF ((x1 = FALSE) AND  ( TRUE )) THEN
        cstate71 := 6; y1 := FALSE; t_start := FALSE;
    END_IF;
END_CASE;

(* Additional processing to handle clocks - in CODESYS, it only starts
    with rising edge and can not be placed inside IF statement *)
IF(t_up = TRUE) THEN
    t_reset := TRUE;
ELSIF(t_start = TRUE AND t_up = FALSE) THEN
    t_up := TRUE;  t_reset := FALSE;
END_IF
t(IN:=t_reset, PT:=T_VALUE);

END_FUNCTION_BLOCK

(* ---- IndustrialAuto8.st ---- *)
FUNCTION_BLOCK FB_G4LTL

   (* Variable definition *)
   VAR_INPUT
      x1	: BOOL;
   END_VAR
   VAR_OUTPUT
      y1	: BOOL;
   END_VAR
   VAR
   (* The total number of states equals to 18 *)
      cstate78	: LINT := 0;
      t0	: TON;
      t0_reset	: BOOL := FALSE;
      t0_up	: BOOL := FALSE;
      t0_start	: BOOL := FALSE;
      t1	: TON;
      t1_reset	: BOOL := FALSE;
      t1_up	: BOOL := FALSE;
      t1_start	: BOOL := FALSE;
   END_VAR

   (* Constant definition (depending on compiler, one might need to move to normal variables) *)

   (* Each time constant has a difference of 1 period (cycle-time); please substract it when needed  *)
   VAR CONST
      T0_VALUE	: TIME := TIME#5s;
      T1_VALUE	: TIME := TIME#3s;
   END_VAR

   (* Control logic *)
CASE cstate78 OF
11:
    IF ((x1 = FALSE) AND  (t0.Q = TRUE) AND  (t1.Q = TRUE)) THEN
        cstate78 := 14; y1 := TRUE; t0_start := FALSE;t1_start := TRUE; t1_up := FALSE;
    ELSIF ((x1 = TRUE) AND  (t0.Q = TRUE) AND  ( TRUE )) THEN
        cstate78 := 10; y1 := FALSE; t0_start := FALSE;t1_start := FALSE;
    ELSIF ((x1 = TRUE) AND  (t0.Q = FALSE) AND  ( TRUE )) THEN
        cstate78 := 11; y1 := FALSE; t0_start := FALSE;t1_start := FALSE;
    ELSIF ((x1 = FALSE) AND  (t0.Q = TRUE) AND  (t1.Q = FALSE)) THEN
        cstate78 := 8; y1 := TRUE; t0_start := FALSE;t1_start := TRUE; t1_up := FALSE;
    ELSIF ((x1 = FALSE) AND  (t0.Q = FALSE) AND  ( TRUE )) THEN
        cstate78 := 1; y1 := FALSE; t0_start := FALSE;t1_start := FALSE;
    END_IF;
12:
    IF ((x1 = TRUE) AND  (t0.Q = TRUE) AND  ( TRUE )) THEN
        cstate78 := 9; y1 := FALSE; t0_start := TRUE; t0_up := FALSE;t1_start := FALSE;
    ELSIF ((x1 = FALSE) AND  ( TRUE ) AND  (t1.Q = FALSE)) THEN
        cstate78 := 16; y1 := FALSE; t0_start := FALSE;t1_start := FALSE;
    ELSIF ((x1 = TRUE) AND  (t0.Q = FALSE) AND  ( TRUE )) THEN
        cstate78 := 3; y1 := FALSE; t0_start := TRUE; t0_up := FALSE;t1_start := FALSE;
    ELSIF ((x1 = FALSE) AND  ( TRUE ) AND  (t1.Q = TRUE)) THEN
        cstate78 := 4; y1 := FALSE; t0_start := FALSE;t1_start := FALSE;
    END_IF;
13:
    IF ((x1 = TRUE) AND  (t0.Q = FALSE) AND  ( TRUE )) THEN
        cstate78 := 3; y1 := FALSE; t0_start := TRUE; t0_up := FALSE;t1_start := FALSE;
    ELSIF ((x1 = TRUE) AND  (t0.Q = TRUE) AND  ( TRUE )) THEN
        cstate78 := 9; y1 := FALSE; t0_start := TRUE; t0_up := FALSE;t1_start := FALSE;
    ELSIF ((x1 = FALSE) AND  ( TRUE ) AND  (t1.Q = TRUE)) THEN
        cstate78 := 4; y1 := FALSE; t0_start := FALSE;t1_start := FALSE;
    ELSIF ((x1 = FALSE) AND  ( TRUE ) AND  (t1.Q = FALSE)) THEN
        cstate78 := 16; y1 := FALSE; t0_start := FALSE;t1_start := FALSE;
    END_IF;
14:
    IF ((x1 = TRUE) AND  (t0.Q = FALSE) AND  (t1.Q = TRUE)) THEN
        cstate78 := 3; y1 := FALSE; t0_start := TRUE; t0_up := FALSE;t1_start := FALSE;
    ELSIF ((x1 = FALSE) AND  ( TRUE ) AND  (t1.Q = TRUE)) THEN
        cstate78 := 12; y1 := FALSE; t0_start := FALSE;t1_start := FALSE;
    ELSIF ((x1 = TRUE) AND  ( TRUE ) AND  (t1.Q = FALSE)) THEN
        cstate78 := 1; y1 := FALSE; t0_start := FALSE;t1_start := FALSE;
    ELSIF ((x1 = FALSE) AND  ( TRUE ) AND  (t1.Q = FALSE)) THEN
        cstate78 := 15; y1 := TRUE; t0_start := FALSE;t1_start := FALSE;
    ELSIF ((x1 = TRUE) AND  (t0.Q = TRUE) AND  (t1.Q = TRUE)) THEN
        cstate78 := 9; y1 := FALSE; t0_start := TRUE; t0_up := FALSE;t1_start := FALSE;
    END_IF;
15:
    IF ((x1 = TRUE) AND  (t0.Q = TRUE) AND  (t1.Q = TRUE)) THEN
        cstate78 := 9; y1 := FALSE; t0_start := TRUE; t0_up := FALSE;t1_start := FALSE;
    ELSIF ((x1 = FALSE) AND  ( TRUE ) AND  (t1.Q = TRUE)) THEN
        cstate78 := 12; y1 := FALSE; t0_start := FALSE;t1_start := FALSE;
    ELSIF ((x1 = TRUE) AND  (t0.Q = FALSE) AND  (t1.Q = TRUE)) THEN
        cstate78 := 3; y1 := FALSE; t0_start := TRUE; t0_up := FALSE;t1_start := FALSE;
    ELSIF ((x1 = TRUE) AND  ( TRUE ) AND  (t1.Q = FALSE)) THEN
        cstate78 := 1; y1 := FALSE; t0_start := FALSE;t1_start := FALSE;
    ELSIF ((x1 = FALSE) AND  ( TRUE ) AND  (t1.Q = FALSE)) THEN
        cstate78 := 15; y1 := TRUE; t0_start := FALSE;t1_start := FALSE;
    END_IF;
16:
    IF ((x1 = TRUE) AND  (t0.Q = TRUE) AND  ( TRUE )) THEN
        cstate78 := 9; y1 := FALSE; t0_start := TRUE; t0_up := FALSE;t1_start := FALSE;
    ELSIF ((x1 = FALSE) AND  ( TRUE ) AND  (t1.Q = TRUE)) THEN
        cstate78 := 4; y1 := FALSE; t0_start := FALSE;t1_start := FALSE;
    ELSIF ((x1 = FALSE) AND  ( TRUE ) AND  (t1.Q = FALSE)) THEN
        cstate78 := 16; y1 := FALSE; t0_start := FALSE;t1_start := FALSE;
    ELSIF ((x1 = TRUE) AND  (t0.Q = FALSE) AND  ( TRUE )) THEN
        cstate78 := 3; y1 := FALSE; t0_start := TRUE; t0_up := FALSE;t1_start := FALSE;
    END_IF;
17:
    IF ((x1 = FALSE) AND  ( TRUE ) AND  (t1.Q = FALSE)) THEN
        cstate78 := 8; y1 := TRUE; t0_start := FALSE;t1_start := TRUE; t1_up := FALSE;
    ELSIF ((x1 = TRUE) AND  (t0.Q = FALSE) AND  ( TRUE )) THEN
        cstate78 := 6; y1 := FALSE; t0_start := FALSE;t1_start := FALSE;
    ELSIF ((x1 = FALSE) AND  ( TRUE ) AND  (t1.Q = TRUE)) THEN
        cstate78 := 14; y1 := TRUE; t0_start := FALSE;t1_start := TRUE; t1_up := FALSE;
    ELSIF ((x1 = TRUE) AND  (t0.Q = TRUE) AND  ( TRUE )) THEN
        cstate78 := 7; y1 := FALSE; t0_start := FALSE;t1_start := FALSE;
    END_IF;
0:
    IF ((x1 = TRUE) AND  (t0.Q = FALSE) AND  ( TRUE )) THEN
        cstate78 := 17; y1 := FALSE; t0_start := FALSE;t1_start := FALSE;
    ELSIF ((x1 = FALSE) AND  ( TRUE ) AND  (t1.Q = FALSE)) THEN
        cstate78 := 2; y1 := FALSE; t0_start := FALSE;t1_start := FALSE;
    ELSIF ((x1 = FALSE) AND  ( TRUE ) AND  (t1.Q = TRUE)) THEN
        cstate78 := 13; y1 := FALSE; t0_start := FALSE;t1_start := FALSE;
    ELSIF ((x1 = TRUE) AND  (t0.Q = TRUE) AND  ( TRUE )) THEN
        cstate78 := 5; y1 := FALSE; t0_start := FALSE;t1_start := FALSE;
    END_IF;
1:
    IF (( TRUE )) THEN
        cstate78 := 1; y1 := FALSE; t0_start := FALSE;t1_start := FALSE;
    END_IF;
2:
    IF ((x1 = TRUE) AND  (t0.Q = FALSE) AND  ( TRUE )) THEN
        cstate78 := 3; y1 := FALSE; t0_start := TRUE; t0_up := FALSE;t1_start := FALSE;
    ELSIF ((x1 = FALSE) AND  ( TRUE ) AND  (t1.Q = FALSE)) THEN
        cstate78 := 16; y1 := FALSE; t0_start := FALSE;t1_start := FALSE;
    ELSIF ((x1 = TRUE) AND  (t0.Q = TRUE) AND  ( TRUE )) THEN
        cstate78 := 9; y1 := FALSE; t0_start := TRUE; t0_up := FALSE;t1_start := FALSE;
    ELSIF ((x1 = FALSE) AND  ( TRUE ) AND  (t1.Q = TRUE)) THEN
        cstate78 := 4; y1 := FALSE; t0_start := FALSE;t1_start := FALSE;
    END_IF;
3:
    IF ((x1 = FALSE) AND  (t0.Q = FALSE) AND  ( TRUE )) THEN
        cstate78 := 1; y1 := FALSE; t0_start := FALSE;t1_start := FALSE;
    ELSIF ((x1 = TRUE) AND  (t0.Q = FALSE) AND  ( TRUE )) THEN
        cstate78 := 11; y1 := FALSE; t0_start := FALSE;t1_start := FALSE;
    ELSIF ((x1 = FALSE) AND  (t0.Q = TRUE) AND  (t1.Q = TRUE)) THEN
        cstate78 := 14; y1 := TRUE; t0_start := FALSE;t1_start := TRUE; t1_up := FALSE;
    ELSIF ((x1 = FALSE) AND  (t0.Q = TRUE) AND  (t1.Q = FALSE)) THEN
        cstate78 := 8; y1 := TRUE; t0_start := FALSE;t1_start := TRUE; t1_up := FALSE;
    ELSIF ((x1 = TRUE) AND  (t0.Q = TRUE) AND  ( TRUE )) THEN
        cstate78 := 10; y1 := FALSE; t0_start := FALSE;t1_start := FALSE;
    END_IF;
4:
    IF ((x1 = FALSE) AND  ( TRUE ) AND  (t1.Q = TRUE)) THEN
        cstate78 := 4; y1 := FALSE; t0_start := FALSE;t1_start := FALSE;
    ELSIF ((x1 = TRUE) AND  (t0.Q = TRUE) AND  ( TRUE )) THEN
        cstate78 := 9; y1 := FALSE; t0_start := TRUE; t0_up := FALSE;t1_start := FALSE;
    ELSIF ((x1 = FALSE) AND  ( TRUE ) AND  (t1.Q = FALSE)) THEN
        cstate78 := 16; y1 := FALSE; t0_start := FALSE;t1_start := FALSE;
    ELSIF ((x1 = TRUE) AND  (t0.Q = FALSE) AND  ( TRUE )) THEN
        cstate78 := 3; y1 := FALSE; t0_start := TRUE; t0_up := FALSE;t1_start := FALSE;
    END_IF;
5:
    IF ((x1 = TRUE) AND  (t0.Q = FALSE) AND  ( TRUE )) THEN
        cstate78 := 6; y1 := FALSE; t0_start := FALSE;t1_start := FALSE;
    ELSIF ((x1 = FALSE) AND  ( TRUE ) AND  (t1.Q = TRUE)) THEN
        cstate78 := 14; y1 := TRUE; t0_start := FALSE;t1_start := TRUE; t1_up := FALSE;
    ELSIF ((x1 = FALSE) AND  ( TRUE ) AND  (t1.Q = FALSE)) THEN
        cstate78 := 8; y1 := TRUE; t0_start := FALSE;t1_start := TRUE; t1_up := FALSE;
    ELSIF ((x1 = TRUE) AND  (t0.Q = TRUE) AND  ( TRUE )) THEN
        cstate78 := 7; y1 := TRUE; t0_start := FALSE;t1_start := FALSE;
    END_IF;
6:
    IF ((x1 = TRUE) AND  (t0.Q = TRUE) AND  ( TRUE )) THEN
        cstate78 := 7; y1 := FALSE; t0_start := FALSE;t1_start := FALSE;
    ELSIF ((x1 = TRUE) AND  (t0.Q = FALSE) AND  ( TRUE )) THEN
        cstate78 := 6; y1 := FALSE; t0_start := FALSE;t1_start := FALSE;
    ELSIF ((x1 = FALSE) AND  ( TRUE ) AND  (t1.Q = TRUE)) THEN
        cstate78 := 14; y1 := TRUE; t0_start := FALSE;t1_start := TRUE; t1_up := FALSE;
    ELSIF ((x1 = FALSE) AND  ( TRUE ) AND  (t1.Q = FALSE)) THEN
        cstate78 := 8; y1 := TRUE; t0_start := FALSE;t1_start := TRUE; t1_up := FALSE;
    END_IF;
7:
    IF ((x1 = FALSE) AND  ( TRUE ) AND  (t1.Q = FALSE)) THEN
        cstate78 := 8; y1 := TRUE; t0_start := FALSE;t1_start := TRUE; t1_up := FALSE;
    ELSIF ((x1 = FALSE) AND  ( TRUE ) AND  (t1.Q = TRUE)) THEN
        cstate78 := 14; y1 := TRUE; t0_start := FALSE;t1_start := TRUE; t1_up := FALSE;
    ELSIF ((x1 = TRUE) AND  (t0.Q = FALSE) AND  ( TRUE )) THEN
        cstate78 := 6; y1 := FALSE; t0_start := FALSE;t1_start := FALSE;
    ELSIF ((x1 = TRUE) AND  (t0.Q = TRUE) AND  ( TRUE )) THEN
        cstate78 := 7; y1 := TRUE; t0_start := FALSE;t1_start := FALSE;
    END_IF;
8:
    IF ((x1 = TRUE) AND  (t0.Q = TRUE) AND  (t1.Q = TRUE)) THEN
        cstate78 := 9; y1 := FALSE; t0_start := TRUE; t0_up := FALSE;t1_start := FALSE;
    ELSIF ((x1 = FALSE) AND  ( TRUE ) AND  (t1.Q = TRUE)) THEN
        cstate78 := 12; y1 := FALSE; t0_start := FALSE;t1_start := FALSE;
    ELSIF ((x1 = TRUE) AND  ( TRUE ) AND  (t1.Q = FALSE)) THEN
        cstate78 := 1; y1 := FALSE; t0_start := FALSE;t1_start := FALSE;
    ELSIF ((x1 = FALSE) AND  ( TRUE ) AND  (t1.Q = FALSE)) THEN
        cstate78 := 15; y1 := TRUE; t0_start := FALSE;t1_start := FALSE;
    ELSIF ((x1 = TRUE) AND  (t0.Q = FALSE) AND  (t1.Q = TRUE)) THEN
        cstate78 := 3; y1 := FALSE; t0_start := TRUE; t0_up := FALSE;t1_start := FALSE;
    END_IF;
9:
    IF ((x1 = TRUE) AND  (t0.Q = TRUE) AND  ( TRUE )) THEN
        cstate78 := 10; y1 := TRUE; t0_start := FALSE;t1_start := FALSE;
    ELSIF ((x1 = FALSE) AND  (t0.Q = FALSE) AND  ( TRUE )) THEN
        cstate78 := 1; y1 := FALSE; t0_start := FALSE;t1_start := FALSE;
    ELSIF ((x1 = FALSE) AND  (t0.Q = TRUE) AND  (t1.Q = TRUE)) THEN
        cstate78 := 14; y1 := TRUE; t0_start := FALSE;t1_start := TRUE; t1_up := FALSE;
    ELSIF ((x1 = TRUE) AND  (t0.Q = FALSE) AND  ( TRUE )) THEN
        cstate78 := 11; y1 := FALSE; t0_start := FALSE;t1_start := FALSE;
    ELSIF ((x1 = FALSE) AND  (t0.Q = TRUE) AND  (t1.Q = FALSE)) THEN
        cstate78 := 8; y1 := TRUE; t0_start := FALSE;t1_start := TRUE; t1_up := FALSE;
    END_IF;
10:
    IF ((x1 = TRUE) AND  (t0.Q = TRUE) AND  ( TRUE )) THEN
        cstate78 := 7; y1 := TRUE; t0_start := FALSE;t1_start := FALSE;
    ELSIF ((x1 = TRUE) AND  (t0.Q = FALSE) AND  ( TRUE )) THEN
        cstate78 := 6; y1 := FALSE; t0_start := FALSE;t1_start := FALSE;
    ELSIF ((x1 = FALSE) AND  ( TRUE ) AND  (t1.Q = TRUE)) THEN
        cstate78 := 14; y1 := TRUE; t0_start := FALSE;t1_start := TRUE; t1_up := FALSE;
    ELSIF ((x1 = FALSE) AND  ( TRUE ) AND  (t1.Q = FALSE)) THEN
        cstate78 := 8; y1 := TRUE; t0_start := FALSE;t1_start := TRUE; t1_up := FALSE;
    END_IF;
END_CASE;

(* Additional processing to handle clocks - in CODESYS, it only starts
    with rising edge and can not be placed inside IF statement *)
IF(t0_up = TRUE) THEN
    t0_reset := TRUE;
ELSIF(t0_start = TRUE AND t0_up = FALSE) THEN
    t0_up := TRUE;  t0_reset := FALSE;
END_IF
t0(IN:=t0_reset, PT:=T0_VALUE);
IF(t1_up = TRUE) THEN
    t1_reset := TRUE;
ELSIF(t1_start = TRUE AND t1_up = FALSE) THEN
    t1_up := TRUE;  t1_reset := FALSE;
END_IF
t1(IN:=t1_reset, PT:=T1_VALUE);

END_FUNCTION_BLOCK

(* ---- Req1.st ---- *)
FUNCTION_BLOCK FB_G4LTL

   (* Variable definition *)
   VAR_INPUT
      req1	: BOOL;
   END_VAR
   VAR_OUTPUT
      grant1	: BOOL;
   END_VAR
   VAR
   (* The total number of states equals to 1 *)
      cstate98	: LINT := 0;
   END_VAR

   (* Control logic *)
CASE cstate98 OF
0:
    IF ((req1 = FALSE)) THEN
        cstate98 := 0; grant1 := FALSE;
    ELSIF ((req1 = TRUE)) THEN
        cstate98 := 0; grant1 := TRUE;
    END_IF;
END_CASE;

END_FUNCTION_BLOCK

(* ---- Req3.st ---- *)
FUNCTION_BLOCK FB_G4LTL

   (* Variable definition *)
   VAR_INPUT
      req	: BOOL;
      cancel	: BOOL;
      go	: BOOL;
   END_VAR
   VAR_OUTPUT
      grant	: BOOL;
   END_VAR
   VAR
   (* The total number of states equals to 22 *)
      cstate23	: LINT := 0;
   END_VAR

   (* Control logic *)
CASE cstate23 OF
11:
    IF ((req = TRUE) AND  (cancel = TRUE) AND  ( TRUE )) THEN
        cstate23 := 8; grant := FALSE;
    ELSIF ((req = TRUE) AND  (cancel = FALSE) AND  ( TRUE )) THEN
        cstate23 := 15; grant := FALSE;
    ELSIF ((req = FALSE) AND  (cancel = FALSE) AND  ( TRUE )) THEN
        cstate23 := 11; grant := FALSE;
    ELSIF ((req = FALSE) AND  (cancel = TRUE) AND  ( TRUE )) THEN
        cstate23 := 19; grant := FALSE;
    END_IF;
12:
    IF ((req = TRUE) AND  (cancel = FALSE) AND  ( TRUE )) THEN
        cstate23 := 13; grant := FALSE;
    ELSIF ((req = FALSE) AND  (cancel = FALSE) AND  ( TRUE )) THEN
        cstate23 := 6; grant := FALSE;
    ELSIF ((req = TRUE) AND  (cancel = TRUE) AND  ( TRUE )) THEN
        cstate23 := 10; grant := FALSE;
    ELSIF ((req = FALSE) AND  (cancel = TRUE) AND  ( TRUE )) THEN
        cstate23 := 20; grant := FALSE;
    END_IF;
13:
    IF ((req = FALSE) AND  (cancel = FALSE) AND  ( TRUE )) THEN
        cstate23 := 7; grant := TRUE;
    ELSIF ((req = TRUE) AND  (cancel = TRUE) AND  ( TRUE )) THEN
        cstate23 := 4; grant := TRUE;
    ELSIF ((req = TRUE) AND  (cancel = FALSE) AND  ( TRUE )) THEN
        cstate23 := 2; grant := TRUE;
    ELSIF ((req = FALSE) AND  (cancel = TRUE) AND  ( TRUE )) THEN
        cstate23 := 18; grant := TRUE;
    END_IF;
14:
    IF ((req = TRUE) AND  (cancel = TRUE) AND  ( TRUE )) THEN
        cstate23 := 4; grant := TRUE;
    ELSIF ((req = TRUE) AND  (cancel = FALSE) AND  ( TRUE )) THEN
        cstate23 := 2; grant := TRUE;
    ELSIF ((req = FALSE) AND  (cancel = TRUE) AND  ( TRUE )) THEN
        cstate23 := 18; grant := TRUE;
    ELSIF ((req = FALSE) AND  (cancel = FALSE) AND  ( TRUE )) THEN
        cstate23 := 7; grant := TRUE;
    END_IF;
15:
    IF ((req = FALSE) AND  (cancel = TRUE) AND  ( TRUE )) THEN
        cstate23 := 9; grant := FALSE;
    ELSIF ((req = TRUE) AND  (cancel = FALSE) AND  ( TRUE )) THEN
        cstate23 := 21; grant := FALSE;
    ELSIF ((req = FALSE) AND  (cancel = FALSE) AND  ( TRUE )) THEN
        cstate23 := 12; grant := FALSE;
    ELSIF ((req = TRUE) AND  (cancel = TRUE) AND  ( TRUE )) THEN
        cstate23 := 17; grant := FALSE;
    END_IF;
16:
    IF (( TRUE )) THEN
        cstate23 := 16; grant := FALSE;
    END_IF;
17:
    IF ((req = FALSE) AND  (cancel = TRUE) AND  (go = TRUE)) THEN
        cstate23 := 1; grant := FALSE;
    ELSIF ((req = TRUE) AND  (cancel = FALSE) AND  (go = TRUE)) THEN
        cstate23 := 3; grant := FALSE;
    ELSIF (( TRUE ) AND  ( TRUE ) AND  (go = FALSE)) THEN
        cstate23 := 16; grant := FALSE;
    ELSIF ((req = FALSE) AND  (cancel = FALSE) AND  (go = TRUE)) THEN
        cstate23 := 14; grant := FALSE;
    ELSIF ((req = TRUE) AND  (cancel = TRUE) AND  (go = TRUE)) THEN
        cstate23 := 5; grant := FALSE;
    END_IF;
18:
    IF ((req = FALSE) AND  (cancel = FALSE) AND  (go = TRUE)) THEN
        cstate23 := 11; grant := FALSE;
    ELSIF ((req = FALSE) AND  (cancel = TRUE) AND  (go = TRUE)) THEN
        cstate23 := 19; grant := FALSE;
    ELSIF (( TRUE ) AND  ( TRUE ) AND  (go = FALSE)) THEN
        cstate23 := 16; grant := FALSE;
    ELSIF ((req = TRUE) AND  (cancel = TRUE) AND  (go = TRUE)) THEN
        cstate23 := 8; grant := FALSE;
    ELSIF ((req = TRUE) AND  (cancel = FALSE) AND  (go = TRUE)) THEN
        cstate23 := 15; grant := FALSE;
    END_IF;
19:
    IF (( TRUE ) AND  ( TRUE ) AND  (go = FALSE)) THEN
        cstate23 := 16; grant := FALSE;
    ELSIF ((req = FALSE) AND  (cancel = TRUE) AND  (go = TRUE)) THEN
        cstate23 := 19; grant := FALSE;
    ELSIF ((req = TRUE) AND  (cancel = FALSE) AND  (go = TRUE)) THEN
        cstate23 := 15; grant := FALSE;
    ELSIF ((req = FALSE) AND  (cancel = FALSE) AND  (go = TRUE)) THEN
        cstate23 := 11; grant := FALSE;
    ELSIF ((req = TRUE) AND  (cancel = TRUE) AND  (go = TRUE)) THEN
        cstate23 := 8; grant := FALSE;
    END_IF;
0:
    IF ((req = FALSE) AND  (cancel = FALSE) AND  ( TRUE )) THEN
        cstate23 := 11; grant := FALSE;
    ELSIF ((req = FALSE) AND  (cancel = TRUE) AND  ( TRUE )) THEN
        cstate23 := 19; grant := FALSE;
    ELSIF ((req = TRUE) AND  (cancel = FALSE) AND  ( TRUE )) THEN
        cstate23 := 15; grant := FALSE;
    ELSIF ((req = TRUE) AND  (cancel = TRUE) AND  ( TRUE )) THEN
        cstate23 := 8; grant := FALSE;
    END_IF;
1:
    IF ((req = TRUE) AND  (cancel = FALSE) AND  (go = TRUE)) THEN
        cstate23 := 2; grant := TRUE;
    ELSIF ((req = FALSE) AND  (cancel = TRUE) AND  (go = TRUE)) THEN
        cstate23 := 18; grant := TRUE;
    ELSIF ((req = FALSE) AND  (cancel = FALSE) AND  (go = TRUE)) THEN
        cstate23 := 7; grant := TRUE;
    ELSIF ((req = TRUE) AND  (cancel = TRUE) AND  (go = TRUE)) THEN
        cstate23 := 4; grant := TRUE;
    ELSIF (( TRUE ) AND  ( TRUE ) AND  (go = FALSE)) THEN
        cstate23 := 16; grant := FALSE;
    END_IF;
2:
    IF ((req = FALSE) AND  (cancel = FALSE) AND  ( TRUE )) THEN
        cstate23 := 12; grant := FALSE;
    ELSIF ((req = TRUE) AND  (cancel = TRUE) AND  ( TRUE )) THEN
        cstate23 := 17; grant := FALSE;
    ELSIF ((req = FALSE) AND  (cancel = TRUE) AND  ( TRUE )) THEN
        cstate23 := 9; grant := FALSE;
    ELSIF ((req = TRUE) AND  (cancel = FALSE) AND  ( TRUE )) THEN
        cstate23 := 21; grant := FALSE;
    END_IF;
3:
    IF ((req = TRUE) AND  (cancel = TRUE) AND  ( TRUE )) THEN
        cstate23 := 4; grant := TRUE;
    ELSIF ((req = FALSE) AND  (cancel = FALSE) AND  ( TRUE )) THEN
        cstate23 := 7; grant := TRUE;
    ELSIF ((req = TRUE) AND  (cancel = FALSE) AND  ( TRUE )) THEN
        cstate23 := 2; grant := TRUE;
    ELSIF ((req = FALSE) AND  (cancel = TRUE) AND  ( TRUE )) THEN
        cstate23 := 18; grant := TRUE;
    END_IF;
4:
    IF (( TRUE ) AND  ( TRUE ) AND  (go = FALSE)) THEN
        cstate23 := 16; grant := FALSE;
    ELSIF ((req = FALSE) AND  (cancel = TRUE) AND  (go = TRUE)) THEN
        cstate23 := 9; grant := FALSE;
    ELSIF ((req = TRUE) AND  (cancel = FALSE) AND  (go = TRUE)) THEN
        cstate23 := 21; grant := FALSE;
    ELSIF ((req = FALSE) AND  (cancel = FALSE) AND  (go = TRUE)) THEN
        cstate23 := 12; grant := FALSE;
    ELSIF ((req = TRUE) AND  (cancel = TRUE) AND  (go = TRUE)) THEN
        cstate23 := 17; grant := FALSE;
    END_IF;
5:
    IF ((req = TRUE) AND  (cancel = FALSE) AND  (go = TRUE)) THEN
        cstate23 := 2; grant := TRUE;
    ELSIF ((req = FALSE) AND  (cancel = TRUE) AND  (go = TRUE)) THEN
        cstate23 := 18; grant := TRUE;
    ELSIF (( TRUE ) AND  ( TRUE ) AND  (go = FALSE)) THEN
        cstate23 := 16; grant := FALSE;
    ELSIF ((req = TRUE) AND  (cancel = TRUE) AND  (go = TRUE)) THEN
        cstate23 := 4; grant := TRUE;
    ELSIF ((req = FALSE) AND  (cancel = FALSE) AND  (go = TRUE)) THEN
        cstate23 := 7; grant := TRUE;
    END_IF;
6:
    IF ((req = FALSE) AND  (cancel = FALSE) AND  ( TRUE )) THEN
        cstate23 := 7; grant := TRUE;
    ELSIF ((req = TRUE) AND  (cancel = TRUE) AND  ( TRUE )) THEN
        cstate23 := 4; grant := TRUE;
    ELSIF ((req = TRUE) AND  (cancel = FALSE) AND  ( TRUE )) THEN
        cstate23 := 2; grant := TRUE;
    ELSIF ((req = FALSE) AND  (cancel = TRUE) AND  ( TRUE )) THEN
        cstate23 := 18; grant := TRUE;
    END_IF;
7:
    IF ((req = TRUE) AND  (cancel = TRUE) AND  ( TRUE )) THEN
        cstate23 := 8; grant := FALSE;
    ELSIF ((req = TRUE) AND  (cancel = FALSE) AND  ( TRUE )) THEN
        cstate23 := 15; grant := FALSE;
    ELSIF ((req = FALSE) AND  (cancel = FALSE) AND  ( TRUE )) THEN
        cstate23 := 11; grant := FALSE;
    ELSIF ((req = FALSE) AND  (cancel = TRUE) AND  ( TRUE )) THEN
        cstate23 := 19; grant := FALSE;
    END_IF;
8:
    IF ((req = FALSE) AND  (cancel = TRUE) AND  (go = TRUE)) THEN
        cstate23 := 9; grant := FALSE;
    ELSIF ((req = TRUE) AND  (cancel = TRUE) AND  (go = TRUE)) THEN
        cstate23 := 17; grant := FALSE;
    ELSIF ((req = FALSE) AND  (cancel = FALSE) AND  (go = TRUE)) THEN
        cstate23 := 12; grant := FALSE;
    ELSIF ((req = TRUE) AND  (cancel = FALSE) AND  (go = TRUE)) THEN
        cstate23 := 21; grant := FALSE;
    ELSIF (( TRUE ) AND  ( TRUE ) AND  (go = FALSE)) THEN
        cstate23 := 16; grant := FALSE;
    END_IF;
9:
    IF ((req = TRUE) AND  (cancel = TRUE) AND  (go = TRUE)) THEN
        cstate23 := 10; grant := FALSE;
    ELSIF ((req = FALSE) AND  (cancel = TRUE) AND  (go = TRUE)) THEN
        cstate23 := 20; grant := FALSE;
    ELSIF ((req = TRUE) AND  (cancel = FALSE) AND  (go = TRUE)) THEN
        cstate23 := 13; grant := FALSE;
    ELSIF (( TRUE ) AND  ( TRUE ) AND  (go = FALSE)) THEN
        cstate23 := 16; grant := FALSE;
    ELSIF ((req = FALSE) AND  (cancel = FALSE) AND  (go = TRUE)) THEN
        cstate23 := 6; grant := FALSE;
    END_IF;
20:
    IF ((req = TRUE) AND  (cancel = FALSE) AND  (go = TRUE)) THEN
        cstate23 := 2; grant := TRUE;
    ELSIF ((req = FALSE) AND  (cancel = TRUE) AND  (go = TRUE)) THEN
        cstate23 := 18; grant := TRUE;
    ELSIF (( TRUE ) AND  ( TRUE ) AND  (go = FALSE)) THEN
        cstate23 := 16; grant := FALSE;
    ELSIF ((req = FALSE) AND  (cancel = FALSE) AND  (go = TRUE)) THEN
        cstate23 := 7; grant := TRUE;
    ELSIF ((req = TRUE) AND  (cancel = TRUE) AND  (go = TRUE)) THEN
        cstate23 := 4; grant := TRUE;
    END_IF;
10:
    IF ((req = FALSE) AND  (cancel = FALSE) AND  (go = TRUE)) THEN
        cstate23 := 7; grant := TRUE;
    ELSIF ((req = TRUE) AND  (cancel = FALSE) AND  (go = TRUE)) THEN
        cstate23 := 2; grant := TRUE;
    ELSIF (( TRUE ) AND  ( TRUE ) AND  (go = FALSE)) THEN
        cstate23 := 16; grant := FALSE;
    ELSIF ((req = FALSE) AND  (cancel = TRUE) AND  (go = TRUE)) THEN
        cstate23 := 18; grant := TRUE;
    ELSIF ((req = TRUE) AND  (cancel = TRUE) AND  (go = TRUE)) THEN
        cstate23 := 4; grant := TRUE;
    END_IF;
21:
    IF ((req = FALSE) AND  (cancel = FALSE) AND  ( TRUE )) THEN
        cstate23 := 14; grant := FALSE;
    ELSIF ((req = TRUE) AND  (cancel = TRUE) AND  ( TRUE )) THEN
        cstate23 := 5; grant := FALSE;
    ELSIF ((req = FALSE) AND  (cancel = TRUE) AND  ( TRUE )) THEN
        cstate23 := 1; grant := FALSE;
    ELSIF ((req = TRUE) AND  (cancel = FALSE) AND  ( TRUE )) THEN
        cstate23 := 3; grant := FALSE;
    END_IF;
END_CASE;

END_FUNCTION_BLOCK

(* ---- Req4.st ---- *)
FUNCTION_BLOCK FB_G4LTL

   (* Variable definition *)
   VAR_INPUT
      req	: BOOL;
      cancel	: BOOL;
      go	: BOOL;
   END_VAR
   VAR_OUTPUT
      grant	: BOOL;
   END_VAR
   VAR
   (* The total number of states equals to 42 *)
      cstate34	: LINT := 0;
   END_VAR

   (* Control logic *)
CASE cstate34 OF
22:
    IF ((req = TRUE) AND  (cancel = FALSE) AND  ( TRUE )) THEN
        cstate34 := 26; grant := FALSE;
    ELSIF ((req = TRUE) AND  (cancel = TRUE) AND  ( TRUE )) THEN
        cstate34 := 14; grant := FALSE;
    ELSIF ((req = FALSE) AND  (cancel = FALSE) AND  ( TRUE )) THEN
        cstate34 := 7; grant := FALSE;
    ELSIF ((req = FALSE) AND  (cancel = TRUE) AND  ( TRUE )) THEN
        cstate34 := 19; grant := FALSE;
    END_IF;
23:
    IF ((req = FALSE) AND  (cancel = TRUE) AND  (go = TRUE)) THEN
        cstate34 := 24; grant := TRUE;
    ELSIF ((req = TRUE) AND  (cancel = FALSE) AND  (go = TRUE)) THEN
        cstate34 := 8; grant := FALSE;
    ELSIF ((req = FALSE) AND  (cancel = FALSE) AND  (go = TRUE)) THEN
        cstate34 := 41; grant := FALSE;
    ELSIF (( TRUE ) AND  ( TRUE ) AND  (go = FALSE)) THEN
        cstate34 := 2; grant := FALSE;
    ELSIF ((req = TRUE) AND  (cancel = TRUE) AND  (go = TRUE)) THEN
        cstate34 := 11; grant := TRUE;
    END_IF;
24:
    IF ((req = TRUE) AND  (cancel = TRUE) AND  (go = TRUE)) THEN
        cstate34 := 18; grant := FALSE;
    ELSIF ((req = TRUE) AND  (cancel = FALSE) AND  (go = TRUE)) THEN
        cstate34 := 22; grant := FALSE;
    ELSIF ((req = FALSE) AND  (cancel = FALSE) AND  (go = TRUE)) THEN
        cstate34 := 32; grant := FALSE;
    ELSIF ((req = FALSE) AND  (cancel = TRUE) AND  (go = TRUE)) THEN
        cstate34 := 17; grant := FALSE;
    ELSIF ((req = FALSE) AND  ( TRUE ) AND  (go = FALSE)) THEN
        cstate34 := 12; grant := FALSE;
    ELSIF ((req = TRUE) AND  ( TRUE ) AND  (go = FALSE)) THEN
        cstate34 := 31; grant := FALSE;
    END_IF;
25:
    IF ((req = FALSE) AND  (cancel = TRUE) AND  ( TRUE )) THEN
        cstate34 := 15; grant := TRUE;
    ELSIF ((req = TRUE) AND  (cancel = FALSE) AND  ( TRUE )) THEN
        cstate34 := 28; grant := TRUE;
    ELSIF ((req = TRUE) AND  (cancel = TRUE) AND  ( TRUE )) THEN
        cstate34 := 9; grant := TRUE;
    ELSIF ((req = FALSE) AND  (cancel = FALSE) AND  ( TRUE )) THEN
        cstate34 := 29; grant := TRUE;
    END_IF;
26:
    IF ((req = TRUE) AND  (cancel = FALSE) AND  ( TRUE )) THEN
        cstate34 := 40; grant := FALSE;
    ELSIF ((req = FALSE) AND  (cancel = FALSE) AND  ( TRUE )) THEN
        cstate34 := 25; grant := FALSE;
    ELSIF ((req = FALSE) AND  (cancel = TRUE) AND  ( TRUE )) THEN
        cstate34 := 15; grant := TRUE;
    ELSIF ((req = TRUE) AND  (cancel = TRUE) AND  ( TRUE )) THEN
        cstate34 := 9; grant := TRUE;
    END_IF;
27:
    IF ((req = FALSE) AND  (cancel = FALSE) AND  (go = TRUE)) THEN
        cstate34 := 25; grant := FALSE;
    ELSIF ((req = FALSE) AND  (cancel = TRUE) AND  (go = TRUE)) THEN
        cstate34 := 15; grant := TRUE;
    ELSIF ((req = FALSE) AND  ( TRUE ) AND  (go = FALSE)) THEN
        cstate34 := 1; grant := FALSE;
    ELSIF ((req = TRUE) AND  (cancel = TRUE) AND  (go = TRUE)) THEN
        cstate34 := 9; grant := TRUE;
    ELSIF ((req = TRUE) AND  (cancel = FALSE) AND  (go = TRUE)) THEN
        cstate34 := 40; grant := FALSE;
    ELSIF ((req = TRUE) AND  ( TRUE ) AND  (go = FALSE)) THEN
        cstate34 := 33; grant := FALSE;
    END_IF;
28:
    IF ((req = TRUE) AND  (cancel = TRUE) AND  ( TRUE )) THEN
        cstate34 := 14; grant := FALSE;
    ELSIF ((req = FALSE) AND  (cancel = FALSE) AND  ( TRUE )) THEN
        cstate34 := 7; grant := FALSE;
    ELSIF ((req = TRUE) AND  (cancel = FALSE) AND  ( TRUE )) THEN
        cstate34 := 26; grant := FALSE;
    ELSIF ((req = FALSE) AND  (cancel = TRUE) AND  ( TRUE )) THEN
        cstate34 := 19; grant := FALSE;
    END_IF;
29:
    IF ((req = FALSE) AND  (cancel = FALSE) AND  ( TRUE )) THEN
        cstate34 := 32; grant := FALSE;
    ELSIF ((req = TRUE) AND  (cancel = TRUE) AND  ( TRUE )) THEN
        cstate34 := 18; grant := FALSE;
    ELSIF ((req = FALSE) AND  (cancel = TRUE) AND  ( TRUE )) THEN
        cstate34 := 17; grant := FALSE;
    ELSIF ((req = TRUE) AND  (cancel = FALSE) AND  ( TRUE )) THEN
        cstate34 := 22; grant := FALSE;
    END_IF;
30:
    IF ((req = TRUE) AND  (cancel = FALSE) AND  (go = TRUE)) THEN
        cstate34 := 6; grant := TRUE;
    ELSIF (( TRUE ) AND  ( TRUE ) AND  (go = FALSE)) THEN
        cstate34 := 2; grant := FALSE;
    ELSIF ((req = TRUE) AND  (cancel = TRUE) AND  (go = TRUE)) THEN
        cstate34 := 11; grant := TRUE;
    ELSIF ((req = FALSE) AND  (cancel = FALSE) AND  (go = TRUE)) THEN
        cstate34 := 5; grant := TRUE;
    ELSIF ((req = FALSE) AND  (cancel = TRUE) AND  (go = TRUE)) THEN
        cstate34 := 24; grant := TRUE;
    END_IF;
31:
    IF (( TRUE ) AND  ( TRUE ) AND  (go = FALSE)) THEN
        cstate34 := 2; grant := FALSE;
    ELSIF ((req = FALSE) AND  (cancel = TRUE) AND  (go = TRUE)) THEN
        cstate34 := 34; grant := FALSE;
    ELSIF ((req = FALSE) AND  (cancel = FALSE) AND  (go = TRUE)) THEN
        cstate34 := 3; grant := FALSE;
    ELSIF ((req = TRUE) AND  (cancel = FALSE) AND  (go = TRUE)) THEN
        cstate34 := 37; grant := FALSE;
    ELSIF ((req = TRUE) AND  (cancel = TRUE) AND  (go = TRUE)) THEN
        cstate34 := 27; grant := FALSE;
    END_IF;
10:
    IF (( TRUE ) AND  ( TRUE ) AND  (go = FALSE)) THEN
        cstate34 := 2; grant := FALSE;
    ELSIF ((req = TRUE) AND  (cancel = FALSE) AND  (go = TRUE)) THEN
        cstate34 := 38; grant := FALSE;
    ELSIF ((req = FALSE) AND  (cancel = FALSE) AND  (go = TRUE)) THEN
        cstate34 := 16; grant := FALSE;
    ELSIF ((req = FALSE) AND  (cancel = TRUE) AND  (go = TRUE)) THEN
        cstate34 := 24; grant := TRUE;
    ELSIF ((req = TRUE) AND  (cancel = TRUE) AND  (go = TRUE)) THEN
        cstate34 := 11; grant := TRUE;
    END_IF;
32:
    IF ((req = FALSE) AND  (cancel = FALSE) AND  ( TRUE )) THEN
        cstate34 := 32; grant := FALSE;
    ELSIF ((req = TRUE) AND  (cancel = FALSE) AND  ( TRUE )) THEN
        cstate34 := 22; grant := FALSE;
    ELSIF ((req = TRUE) AND  (cancel = TRUE) AND  ( TRUE )) THEN
        cstate34 := 18; grant := FALSE;
    ELSIF ((req = FALSE) AND  (cancel = TRUE) AND  ( TRUE )) THEN
        cstate34 := 17; grant := FALSE;
    END_IF;
11:
    IF ((req = TRUE) AND  ( TRUE ) AND  (go = FALSE)) THEN
        cstate34 := 10; grant := FALSE;
    ELSIF ((req = TRUE) AND  (cancel = FALSE) AND  (go = TRUE)) THEN
        cstate34 := 26; grant := FALSE;
    ELSIF ((req = FALSE) AND  (cancel = FALSE) AND  (go = TRUE)) THEN
        cstate34 := 7; grant := FALSE;
    ELSIF ((req = TRUE) AND  (cancel = TRUE) AND  (go = TRUE)) THEN
        cstate34 := 14; grant := FALSE;
    ELSIF ((req = FALSE) AND  (cancel = TRUE) AND  (go = TRUE)) THEN
        cstate34 := 19; grant := FALSE;
    ELSIF ((req = FALSE) AND  ( TRUE ) AND  (go = FALSE)) THEN
        cstate34 := 23; grant := FALSE;
    END_IF;
33:
    IF ((req = FALSE) AND  (cancel = FALSE) AND  (go = TRUE)) THEN
        cstate34 := 5; grant := TRUE;
    ELSIF ((req = TRUE) AND  (cancel = FALSE) AND  (go = TRUE)) THEN
        cstate34 := 6; grant := TRUE;
    ELSIF ((req = FALSE) AND  (cancel = TRUE) AND  (go = TRUE)) THEN
        cstate34 := 24; grant := TRUE;
    ELSIF (( TRUE ) AND  ( TRUE ) AND  (go = FALSE)) THEN
        cstate34 := 2; grant := FALSE;
    ELSIF ((req = TRUE) AND  (cancel = TRUE) AND  (go = TRUE)) THEN
        cstate34 := 11; grant := TRUE;
    END_IF;
12:
    IF ((req = FALSE) AND  (cancel = TRUE) AND  (go = TRUE)) THEN
        cstate34 := 13; grant := FALSE;
    ELSIF ((req = TRUE) AND  (cancel = FALSE) AND  (go = TRUE)) THEN
        cstate34 := 35; grant := FALSE;
    ELSIF (( TRUE ) AND  ( TRUE ) AND  (go = FALSE)) THEN
        cstate34 := 2; grant := FALSE;
    ELSIF ((req = TRUE) AND  (cancel = TRUE) AND  (go = TRUE)) THEN
        cstate34 := 39; grant := FALSE;
    ELSIF ((req = FALSE) AND  (cancel = FALSE) AND  (go = TRUE)) THEN
        cstate34 := 21; grant := FALSE;
    END_IF;
34:
    IF ((req = TRUE) AND  (cancel = TRUE) AND  (go = TRUE)) THEN
        cstate34 := 9; grant := TRUE;
    ELSIF ((req = FALSE) AND  ( TRUE ) AND  (go = FALSE)) THEN
        cstate34 := 30; grant := FALSE;
    ELSIF ((req = FALSE) AND  (cancel = TRUE) AND  (go = TRUE)) THEN
        cstate34 := 15; grant := TRUE;
    ELSIF ((req = TRUE) AND  ( TRUE ) AND  (go = FALSE)) THEN
        cstate34 := 20; grant := FALSE;
    ELSIF ((req = TRUE) AND  (cancel = FALSE) AND  (go = TRUE)) THEN
        cstate34 := 36; grant := FALSE;
    ELSIF ((req = FALSE) AND  (cancel = FALSE) AND  (go = TRUE)) THEN
        cstate34 := 4; grant := FALSE;
    END_IF;
13:
    IF ((req = FALSE) AND  (cancel = FALSE) AND  (go = TRUE)) THEN
        cstate34 := 32; grant := FALSE;
    ELSIF ((req = FALSE) AND  ( TRUE ) AND  (go = FALSE)) THEN
        cstate34 := 12; grant := FALSE;
    ELSIF ((req = TRUE) AND  (cancel = TRUE) AND  (go = TRUE)) THEN
        cstate34 := 18; grant := FALSE;
    ELSIF ((req = FALSE) AND  (cancel = TRUE) AND  (go = TRUE)) THEN
        cstate34 := 17; grant := FALSE;
    ELSIF ((req = TRUE) AND  ( TRUE ) AND  (go = FALSE)) THEN
        cstate34 := 31; grant := FALSE;
    ELSIF ((req = TRUE) AND  (cancel = FALSE) AND  (go = TRUE)) THEN
        cstate34 := 22; grant := FALSE;
    END_IF;
35:
    IF ((req = TRUE) AND  (cancel = FALSE) AND  ( TRUE )) THEN
        cstate34 := 26; grant := FALSE;
    ELSIF ((req = FALSE) AND  (cancel = FALSE) AND  ( TRUE )) THEN
        cstate34 := 7; grant := FALSE;
    ELSIF ((req = TRUE) AND  (cancel = TRUE) AND  ( TRUE )) THEN
        cstate34 := 14; grant := FALSE;
    ELSIF ((req = FALSE) AND  (cancel = TRUE) AND  ( TRUE )) THEN
        cstate34 := 19; grant := FALSE;
    END_IF;
14:
    IF ((req = FALSE) AND  (cancel = TRUE) AND  (go = TRUE)) THEN
        cstate34 := 15; grant := TRUE;
    ELSIF ((req = FALSE) AND  ( TRUE ) AND  (go = FALSE)) THEN
        cstate34 := 1; grant := FALSE;
    ELSIF ((req = TRUE) AND  ( TRUE ) AND  (go = FALSE)) THEN
        cstate34 := 33; grant := FALSE;
    ELSIF ((req = TRUE) AND  (cancel = TRUE) AND  (go = TRUE)) THEN
        cstate34 := 9; grant := TRUE;
    ELSIF ((req = TRUE) AND  (cancel = FALSE) AND  (go = TRUE)) THEN
        cstate34 := 40; grant := FALSE;
    ELSIF ((req = FALSE) AND  (cancel = FALSE) AND  (go = TRUE)) THEN
        cstate34 := 25; grant := FALSE;
    END_IF;
36:
    IF ((req = TRUE) AND  (cancel = TRUE) AND  ( TRUE )) THEN
        cstate34 := 9; grant := TRUE;
    ELSIF ((req = FALSE) AND  (cancel = TRUE) AND  ( TRUE )) THEN
        cstate34 := 15; grant := TRUE;
    ELSIF ((req = TRUE) AND  (cancel = FALSE) AND  ( TRUE )) THEN
        cstate34 := 28; grant := TRUE;
    ELSIF ((req = FALSE) AND  (cancel = FALSE) AND  ( TRUE )) THEN
        cstate34 := 29; grant := TRUE;
    END_IF;
15:
    IF ((req = TRUE) AND  (cancel = TRUE) AND  (go = TRUE)) THEN
        cstate34 := 18; grant := FALSE;
    ELSIF ((req = TRUE) AND  (cancel = FALSE) AND  (go = TRUE)) THEN
        cstate34 := 22; grant := FALSE;
    ELSIF ((req = FALSE) AND  (cancel = TRUE) AND  (go = TRUE)) THEN
        cstate34 := 17; grant := FALSE;
    ELSIF ((req = TRUE) AND  ( TRUE ) AND  (go = FALSE)) THEN
        cstate34 := 31; grant := FALSE;
    ELSIF ((req = FALSE) AND  ( TRUE ) AND  (go = FALSE)) THEN
        cstate34 := 12; grant := FALSE;
    ELSIF ((req = FALSE) AND  (cancel = FALSE) AND  (go = TRUE)) THEN
        cstate34 := 32; grant := FALSE;
    END_IF;
37:
    IF ((req = TRUE) AND  (cancel = TRUE) AND  ( TRUE )) THEN
        cstate34 := 9; grant := TRUE;
    ELSIF ((req = FALSE) AND  (cancel = FALSE) AND  ( TRUE )) THEN
        cstate34 := 25; grant := FALSE;
    ELSIF ((req = FALSE) AND  (cancel = TRUE) AND  ( TRUE )) THEN
        cstate34 := 15; grant := TRUE;
    ELSIF ((req = TRUE) AND  (cancel = FALSE) AND  ( TRUE )) THEN
        cstate34 := 40; grant := FALSE;
    END_IF;
16:
    IF ((req = TRUE) AND  (cancel = TRUE) AND  ( TRUE )) THEN
        cstate34 := 9; grant := TRUE;
    ELSIF ((req = FALSE) AND  (cancel = FALSE) AND  ( TRUE )) THEN
        cstate34 := 29; grant := TRUE;
    ELSIF ((req = TRUE) AND  (cancel = FALSE) AND  ( TRUE )) THEN
        cstate34 := 28; grant := TRUE;
    ELSIF ((req = FALSE) AND  (cancel = TRUE) AND  ( TRUE )) THEN
        cstate34 := 15; grant := TRUE;
    END_IF;
38:
    IF ((req = FALSE) AND  (cancel = FALSE) AND  ( TRUE )) THEN
        cstate34 := 29; grant := TRUE;
    ELSIF ((req = TRUE) AND  (cancel = FALSE) AND  ( TRUE )) THEN
        cstate34 := 28; grant := TRUE;
    ELSIF ((req = TRUE) AND  (cancel = TRUE) AND  ( TRUE )) THEN
        cstate34 := 9; grant := TRUE;
    ELSIF ((req = FALSE) AND  (cancel = TRUE) AND  ( TRUE )) THEN
        cstate34 := 15; grant := TRUE;
    END_IF;
17:
    IF ((req = FALSE) AND  ( TRUE ) AND  (go = FALSE)) THEN
        cstate34 := 12; grant := FALSE;
    ELSIF ((req = FALSE) AND  (cancel = TRUE) AND  (go = TRUE)) THEN
        cstate34 := 17; grant := FALSE;
    ELSIF ((req = TRUE) AND  (cancel = TRUE) AND  (go = TRUE)) THEN
        cstate34 := 18; grant := FALSE;
    ELSIF ((req = TRUE) AND  ( TRUE ) AND  (go = FALSE)) THEN
        cstate34 := 31; grant := FALSE;
    ELSIF ((req = FALSE) AND  (cancel = FALSE) AND  (go = TRUE)) THEN
        cstate34 := 32; grant := FALSE;
    ELSIF ((req = TRUE) AND  (cancel = FALSE) AND  (go = TRUE)) THEN
        cstate34 := 22; grant := FALSE;
    END_IF;
39:
    IF ((req = FALSE) AND  (cancel = TRUE) AND  (go = TRUE)) THEN
        cstate34 := 19; grant := FALSE;
    ELSIF ((req = FALSE) AND  ( TRUE ) AND  (go = FALSE)) THEN
        cstate34 := 23; grant := FALSE;
    ELSIF ((req = TRUE) AND  ( TRUE ) AND  (go = FALSE)) THEN
        cstate34 := 10; grant := FALSE;
    ELSIF ((req = TRUE) AND  (cancel = TRUE) AND  (go = TRUE)) THEN
        cstate34 := 14; grant := FALSE;
    ELSIF ((req = TRUE) AND  (cancel = FALSE) AND  (go = TRUE)) THEN
        cstate34 := 26; grant := FALSE;
    ELSIF ((req = FALSE) AND  (cancel = FALSE) AND  (go = TRUE)) THEN
        cstate34 := 7; grant := FALSE;
    END_IF;
18:
    IF ((req = TRUE) AND  ( TRUE ) AND  (go = FALSE)) THEN
        cstate34 := 10; grant := FALSE;
    ELSIF ((req = FALSE) AND  (cancel = TRUE) AND  (go = TRUE)) THEN
        cstate34 := 19; grant := FALSE;
    ELSIF ((req = FALSE) AND  ( TRUE ) AND  (go = FALSE)) THEN
        cstate34 := 23; grant := FALSE;
    ELSIF ((req = TRUE) AND  (cancel = TRUE) AND  (go = TRUE)) THEN
        cstate34 := 14; grant := FALSE;
    ELSIF ((req = TRUE) AND  (cancel = FALSE) AND  (go = TRUE)) THEN
        cstate34 := 26; grant := FALSE;
    ELSIF ((req = FALSE) AND  (cancel = FALSE) AND  (go = TRUE)) THEN
        cstate34 := 7; grant := FALSE;
    END_IF;
19:
    IF ((req = TRUE) AND  ( TRUE ) AND  (go = FALSE)) THEN
        cstate34 := 20; grant := FALSE;
    ELSIF ((req = TRUE) AND  (cancel = TRUE) AND  (go = TRUE)) THEN
        cstate34 := 9; grant := TRUE;
    ELSIF ((req = FALSE) AND  (cancel = TRUE) AND  (go = TRUE)) THEN
        cstate34 := 15; grant := TRUE;
    ELSIF ((req = FALSE) AND  ( TRUE ) AND  (go = FALSE)) THEN
        cstate34 := 30; grant := FALSE;
    ELSIF ((req = TRUE) AND  (cancel = FALSE) AND  (go = TRUE)) THEN
        cstate34 := 36; grant := FALSE;
    ELSIF ((req = FALSE) AND  (cancel = FALSE) AND  (go = TRUE)) THEN
        cstate34 := 4; grant := FALSE;
    END_IF;
0:
    IF ((req = TRUE) AND  (cancel = FALSE) AND  ( TRUE )) THEN
        cstate34 := 35; grant := FALSE;
    ELSIF ((req = FALSE) AND  (cancel = TRUE) AND  ( TRUE )) THEN
        cstate34 := 13; grant := FALSE;
    ELSIF ((req = TRUE) AND  (cancel = TRUE) AND  ( TRUE )) THEN
        cstate34 := 39; grant := FALSE;
    ELSIF ((req = FALSE) AND  (cancel = FALSE) AND  ( TRUE )) THEN
        cstate34 := 21; grant := FALSE;
    END_IF;
1:
    IF (( TRUE ) AND  ( TRUE ) AND  (go = FALSE)) THEN
        cstate34 := 2; grant := FALSE;
    ELSIF ((req = FALSE) AND  (cancel = FALSE) AND  (go = TRUE)) THEN
        cstate34 := 5; grant := TRUE;
    ELSIF ((req = FALSE) AND  (cancel = TRUE) AND  (go = TRUE)) THEN
        cstate34 := 24; grant := TRUE;
    ELSIF ((req = TRUE) AND  (cancel = TRUE) AND  (go = TRUE)) THEN
        cstate34 := 11; grant := TRUE;
    ELSIF ((req = TRUE) AND  (cancel = FALSE) AND  (go = TRUE)) THEN
        cstate34 := 6; grant := TRUE;
    END_IF;
2:
    IF (( TRUE )) THEN
        cstate34 := 2; grant := FALSE;
    END_IF;
3:
    IF ((req = FALSE) AND  (cancel = FALSE) AND  ( TRUE )) THEN
        cstate34 := 4; grant := FALSE;
    ELSIF ((req = TRUE) AND  (cancel = TRUE) AND  ( TRUE )) THEN
        cstate34 := 9; grant := TRUE;
    ELSIF ((req = TRUE) AND  (cancel = FALSE) AND  ( TRUE )) THEN
        cstate34 := 36; grant := FALSE;
    ELSIF ((req = FALSE) AND  (cancel = TRUE) AND  ( TRUE )) THEN
        cstate34 := 15; grant := TRUE;
    END_IF;
4:
    IF ((req = TRUE) AND  (cancel = FALSE) AND  ( TRUE )) THEN
        cstate34 := 28; grant := TRUE;
    ELSIF ((req = FALSE) AND  (cancel = FALSE) AND  ( TRUE )) THEN
        cstate34 := 29; grant := TRUE;
    ELSIF ((req = FALSE) AND  (cancel = TRUE) AND  ( TRUE )) THEN
        cstate34 := 15; grant := TRUE;
    ELSIF ((req = TRUE) AND  (cancel = TRUE) AND  ( TRUE )) THEN
        cstate34 := 9; grant := TRUE;
    END_IF;
5:
    IF ((req = FALSE) AND  (cancel = TRUE) AND  ( TRUE )) THEN
        cstate34 := 17; grant := FALSE;
    ELSIF ((req = FALSE) AND  (cancel = FALSE) AND  ( TRUE )) THEN
        cstate34 := 32; grant := FALSE;
    ELSIF ((req = TRUE) AND  (cancel = TRUE) AND  ( TRUE )) THEN
        cstate34 := 18; grant := FALSE;
    ELSIF ((req = TRUE) AND  (cancel = FALSE) AND  ( TRUE )) THEN
        cstate34 := 22; grant := FALSE;
    END_IF;
6:
    IF ((req = FALSE) AND  (cancel = FALSE) AND  ( TRUE )) THEN
        cstate34 := 7; grant := FALSE;
    ELSIF ((req = FALSE) AND  (cancel = TRUE) AND  ( TRUE )) THEN
        cstate34 := 19; grant := FALSE;
    ELSIF ((req = TRUE) AND  (cancel = FALSE) AND  ( TRUE )) THEN
        cstate34 := 26; grant := FALSE;
    ELSIF ((req = TRUE) AND  (cancel = TRUE) AND  ( TRUE )) THEN
        cstate34 := 14; grant := FALSE;
    END_IF;
7:
    IF ((req = TRUE) AND  (cancel = TRUE) AND  ( TRUE )) THEN
        cstate34 := 9; grant := TRUE;
    ELSIF ((req = FALSE) AND  (cancel = FALSE) AND  ( TRUE )) THEN
        cstate34 := 4; grant := FALSE;
    ELSIF ((req = TRUE) AND  (cancel = FALSE) AND  ( TRUE )) THEN
        cstate34 := 36; grant := FALSE;
    ELSIF ((req = FALSE) AND  (cancel = TRUE) AND  ( TRUE )) THEN
        cstate34 := 15; grant := TRUE;
    END_IF;
8:
    IF ((req = TRUE) AND  (cancel = TRUE) AND  ( TRUE )) THEN
        cstate34 := 9; grant := TRUE;
    ELSIF ((req = FALSE) AND  (cancel = FALSE) AND  ( TRUE )) THEN
        cstate34 := 29; grant := TRUE;
    ELSIF ((req = FALSE) AND  (cancel = TRUE) AND  ( TRUE )) THEN
        cstate34 := 15; grant := TRUE;
    ELSIF ((req = TRUE) AND  (cancel = FALSE) AND  ( TRUE )) THEN
        cstate34 := 28; grant := TRUE;
    END_IF;
9:
    IF ((req = FALSE) AND  (cancel = FALSE) AND  (go = TRUE)) THEN
        cstate34 := 7; grant := FALSE;
    ELSIF ((req = TRUE) AND  (cancel = FALSE) AND  (go = TRUE)) THEN
        cstate34 := 26; grant := FALSE;
    ELSIF ((req = TRUE) AND  ( TRUE ) AND  (go = FALSE)) THEN
        cstate34 := 10; grant := FALSE;
    ELSIF ((req = TRUE) AND  (cancel = TRUE) AND  (go = TRUE)) THEN
        cstate34 := 14; grant := FALSE;
    ELSIF ((req = FALSE) AND  (cancel = TRUE) AND  (go = TRUE)) THEN
        cstate34 := 19; grant := FALSE;
    ELSIF ((req = FALSE) AND  ( TRUE ) AND  (go = FALSE)) THEN
        cstate34 := 23; grant := FALSE;
    END_IF;
40:
    IF ((req = TRUE) AND  (cancel = FALSE) AND  ( TRUE )) THEN
        cstate34 := 28; grant := TRUE;
    ELSIF ((req = FALSE) AND  (cancel = FALSE) AND  ( TRUE )) THEN
        cstate34 := 29; grant := TRUE;
    ELSIF ((req = TRUE) AND  (cancel = TRUE) AND  ( TRUE )) THEN
        cstate34 := 9; grant := TRUE;
    ELSIF ((req = FALSE) AND  (cancel = TRUE) AND  ( TRUE )) THEN
        cstate34 := 15; grant := TRUE;
    END_IF;
41:
    IF ((req = FALSE) AND  (cancel = FALSE) AND  ( TRUE )) THEN
        cstate34 := 29; grant := TRUE;
    ELSIF ((req = TRUE) AND  (cancel = FALSE) AND  ( TRUE )) THEN
        cstate34 := 28; grant := TRUE;
    ELSIF ((req = TRUE) AND  (cancel = TRUE) AND  ( TRUE )) THEN
        cstate34 := 9; grant := TRUE;
    ELSIF ((req = FALSE) AND  (cancel = TRUE) AND  ( TRUE )) THEN
        cstate34 := 15; grant := TRUE;
    END_IF;
20:
    IF ((req = FALSE) AND  (cancel = FALSE) AND  (go = TRUE)) THEN
        cstate34 := 5; grant := TRUE;
    ELSIF (( TRUE ) AND  ( TRUE ) AND  (go = FALSE)) THEN
        cstate34 := 2; grant := FALSE;
    ELSIF ((req = TRUE) AND  (cancel = FALSE) AND  (go = TRUE)) THEN
        cstate34 := 6; grant := TRUE;
    ELSIF ((req = FALSE) AND  (cancel = TRUE) AND  (go = TRUE)) THEN
        cstate34 := 24; grant := TRUE;
    ELSIF ((req = TRUE) AND  (cancel = TRUE) AND  (go = TRUE)) THEN
        cstate34 := 11; grant := TRUE;
    END_IF;
21:
    IF ((req = TRUE) AND  (cancel = FALSE) AND  ( TRUE )) THEN
        cstate34 := 22; grant := FALSE;
    ELSIF ((req = TRUE) AND  (cancel = TRUE) AND  ( TRUE )) THEN
        cstate34 := 18; grant := FALSE;
    ELSIF ((req = FALSE) AND  (cancel = FALSE) AND  ( TRUE )) THEN
        cstate34 := 32; grant := FALSE;
    ELSIF ((req = FALSE) AND  (cancel = TRUE) AND  ( TRUE )) THEN
        cstate34 := 17; grant := FALSE;
    END_IF;
END_CASE;

END_FUNCTION_BLOCK

(* ---- Req5.st ---- *)
FUNCTION_BLOCK FB_G4LTL

   (* Variable definition *)
   VAR_INPUT
      req	: BOOL;
      cancel	: BOOL;
      go	: BOOL;
   END_VAR
   VAR_OUTPUT
      grant	: BOOL;
   END_VAR
   VAR
   (* The total number of states equals to 28 *)
      cstate52	: LINT := 0;
   END_VAR

   (* Control logic *)
CASE cstate52 OF
22:
    IF (( TRUE )) THEN
        cstate52 := 22; grant := FALSE;
    END_IF;
23:
    IF ((req = TRUE) AND  (cancel = FALSE) AND  ( TRUE )) THEN
        cstate52 := 24; grant := FALSE;
    ELSIF ((req = FALSE) AND  (cancel = TRUE) AND  ( TRUE )) THEN
        cstate52 := 2; grant := FALSE;
    ELSIF ((req = FALSE) AND  (cancel = FALSE) AND  ( TRUE )) THEN
        cstate52 := 5; grant := FALSE;
    ELSIF ((req = TRUE) AND  (cancel = TRUE) AND  ( TRUE )) THEN
        cstate52 := 6; grant := FALSE;
    END_IF;
24:
    IF ((req = TRUE) AND  (cancel = TRUE) AND  ( TRUE )) THEN
        cstate52 := 6; grant := FALSE;
    ELSIF ((req = FALSE) AND  (cancel = FALSE) AND  ( TRUE )) THEN
        cstate52 := 18; grant := TRUE;
    ELSIF ((req = FALSE) AND  (cancel = TRUE) AND  ( TRUE )) THEN
        cstate52 := 2; grant := FALSE;
    ELSIF ((req = TRUE) AND  (cancel = FALSE) AND  ( TRUE )) THEN
        cstate52 := 8; grant := TRUE;
    END_IF;
25:
    IF ((req = FALSE) AND  (cancel = TRUE) AND  ( TRUE )) THEN
        cstate52 := 2; grant := FALSE;
    ELSIF ((req = TRUE) AND  (cancel = FALSE) AND  ( TRUE )) THEN
        cstate52 := 1; grant := FALSE;
    ELSIF ((req = TRUE) AND  (cancel = TRUE) AND  ( TRUE )) THEN
        cstate52 := 6; grant := FALSE;
    ELSIF ((req = FALSE) AND  (cancel = FALSE) AND  ( TRUE )) THEN
        cstate52 := 9; grant := FALSE;
    END_IF;
26:
    IF ((req = TRUE) AND  (cancel = FALSE) AND  ( TRUE )) THEN
        cstate52 := 8; grant := TRUE;
    ELSIF ((req = TRUE) AND  (cancel = TRUE) AND  ( TRUE )) THEN
        cstate52 := 6; grant := FALSE;
    ELSIF ((req = FALSE) AND  (cancel = FALSE) AND  ( TRUE )) THEN
        cstate52 := 18; grant := TRUE;
    ELSIF ((req = FALSE) AND  (cancel = TRUE) AND  ( TRUE )) THEN
        cstate52 := 2; grant := FALSE;
    END_IF;
27:
    IF ((req = TRUE) AND  (cancel = FALSE) AND  (go = TRUE)) THEN
        cstate52 := 26; grant := FALSE;
    ELSIF (( TRUE ) AND  ( TRUE ) AND  (go = FALSE)) THEN
        cstate52 := 22; grant := FALSE;
    ELSIF ((req = TRUE) AND  (cancel = TRUE) AND  (go = TRUE)) THEN
        cstate52 := 16; grant := FALSE;
    ELSIF ((req = FALSE) AND  (cancel = FALSE) AND  (go = TRUE)) THEN
        cstate52 := 15; grant := FALSE;
    ELSIF ((req = FALSE) AND  (cancel = TRUE) AND  (go = TRUE)) THEN
        cstate52 := 20; grant := FALSE;
    END_IF;
10:
    IF ((req = FALSE) AND  (cancel = FALSE) AND  (go = TRUE)) THEN
        cstate52 := 11; grant := FALSE;
    ELSIF ((req = TRUE) AND  (cancel = FALSE) AND  (go = TRUE)) THEN
        cstate52 := 17; grant := FALSE;
    ELSIF (( TRUE ) AND  ( TRUE ) AND  (go = FALSE)) THEN
        cstate52 := 22; grant := FALSE;
    ELSIF ((req = FALSE) AND  (cancel = TRUE) AND  (go = TRUE)) THEN
        cstate52 := 20; grant := FALSE;
    ELSIF ((req = TRUE) AND  (cancel = TRUE) AND  (go = TRUE)) THEN
        cstate52 := 16; grant := FALSE;
    END_IF;
11:
    IF ((req = TRUE) AND  (cancel = FALSE) AND  ( TRUE )) THEN
        cstate52 := 8; grant := TRUE;
    ELSIF ((req = FALSE) AND  (cancel = TRUE) AND  ( TRUE )) THEN
        cstate52 := 2; grant := FALSE;
    ELSIF ((req = FALSE) AND  (cancel = FALSE) AND  ( TRUE )) THEN
        cstate52 := 18; grant := TRUE;
    ELSIF ((req = TRUE) AND  (cancel = TRUE) AND  ( TRUE )) THEN
        cstate52 := 6; grant := FALSE;
    END_IF;
12:
    IF ((req = FALSE) AND  (cancel = FALSE) AND  ( TRUE )) THEN
        cstate52 := 13; grant := FALSE;
    ELSIF ((req = TRUE) AND  (cancel = TRUE) AND  ( TRUE )) THEN
        cstate52 := 6; grant := FALSE;
    ELSIF ((req = TRUE) AND  (cancel = FALSE) AND  ( TRUE )) THEN
        cstate52 := 19; grant := FALSE;
    ELSIF ((req = FALSE) AND  (cancel = TRUE) AND  ( TRUE )) THEN
        cstate52 := 2; grant := FALSE;
    END_IF;
13:
    IF ((req = TRUE) AND  (cancel = FALSE) AND  ( TRUE )) THEN
        cstate52 := 8; grant := TRUE;
    ELSIF ((req = FALSE) AND  (cancel = FALSE) AND  ( TRUE )) THEN
        cstate52 := 18; grant := TRUE;
    ELSIF ((req = TRUE) AND  (cancel = TRUE) AND  ( TRUE )) THEN
        cstate52 := 6; grant := FALSE;
    ELSIF ((req = FALSE) AND  (cancel = TRUE) AND  ( TRUE )) THEN
        cstate52 := 2; grant := FALSE;
    END_IF;
14:
    IF ((req = TRUE) AND  (cancel = TRUE) AND  ( TRUE )) THEN
        cstate52 := 6; grant := FALSE;
    ELSIF ((req = FALSE) AND  (cancel = TRUE) AND  ( TRUE )) THEN
        cstate52 := 2; grant := FALSE;
    ELSIF ((req = TRUE) AND  (cancel = FALSE) AND  ( TRUE )) THEN
        cstate52 := 19; grant := FALSE;
    ELSIF ((req = FALSE) AND  (cancel = FALSE) AND  ( TRUE )) THEN
        cstate52 := 13; grant := FALSE;
    END_IF;
15:
    IF ((req = FALSE) AND  (cancel = TRUE) AND  ( TRUE )) THEN
        cstate52 := 2; grant := FALSE;
    ELSIF ((req = TRUE) AND  (cancel = FALSE) AND  ( TRUE )) THEN
        cstate52 := 8; grant := TRUE;
    ELSIF ((req = FALSE) AND  (cancel = FALSE) AND  ( TRUE )) THEN
        cstate52 := 18; grant := TRUE;
    ELSIF ((req = TRUE) AND  (cancel = TRUE) AND  ( TRUE )) THEN
        cstate52 := 6; grant := FALSE;
    END_IF;
16:
    IF ((req = TRUE) AND  (cancel = FALSE) AND  (go = FALSE)) THEN
        cstate52 := 10; grant := FALSE;
    ELSIF ((req = FALSE) AND  (cancel = FALSE) AND  (go = TRUE)) THEN
        cstate52 := 7; grant := FALSE;
    ELSIF ((req = TRUE) AND  (cancel = TRUE) AND  (go = TRUE)) THEN
        cstate52 := 6; grant := FALSE;
    ELSIF ((req = FALSE) AND  (cancel = TRUE) AND  (go = FALSE)) THEN
        cstate52 := 3; grant := FALSE;
    ELSIF ((req = FALSE) AND  (cancel = TRUE) AND  (go = TRUE)) THEN
        cstate52 := 2; grant := FALSE;
    ELSIF ((req = FALSE) AND  (cancel = FALSE) AND  (go = FALSE)) THEN
        cstate52 := 27; grant := FALSE;
    ELSIF ((req = TRUE) AND  (cancel = TRUE) AND  (go = FALSE)) THEN
        cstate52 := 21; grant := FALSE;
    ELSIF ((req = TRUE) AND  (cancel = FALSE) AND  (go = TRUE)) THEN
        cstate52 := 12; grant := FALSE;
    END_IF;
17:
    IF ((req = FALSE) AND  (cancel = FALSE) AND  ( TRUE )) THEN
        cstate52 := 18; grant := TRUE;
    ELSIF ((req = TRUE) AND  (cancel = FALSE) AND  ( TRUE )) THEN
        cstate52 := 8; grant := TRUE;
    ELSIF ((req = TRUE) AND  (cancel = TRUE) AND  ( TRUE )) THEN
        cstate52 := 6; grant := FALSE;
    ELSIF ((req = FALSE) AND  (cancel = TRUE) AND  ( TRUE )) THEN
        cstate52 := 2; grant := FALSE;
    END_IF;
18:
    IF ((req = FALSE) AND  (cancel = TRUE) AND  ( TRUE )) THEN
        cstate52 := 2; grant := FALSE;
    ELSIF ((req = FALSE) AND  (cancel = FALSE) AND  ( TRUE )) THEN
        cstate52 := 9; grant := FALSE;
    ELSIF ((req = TRUE) AND  (cancel = FALSE) AND  ( TRUE )) THEN
        cstate52 := 1; grant := FALSE;
    ELSIF ((req = TRUE) AND  (cancel = TRUE) AND  ( TRUE )) THEN
        cstate52 := 6; grant := FALSE;
    END_IF;
19:
    IF ((req = FALSE) AND  (cancel = FALSE) AND  ( TRUE )) THEN
        cstate52 := 18; grant := TRUE;
    ELSIF ((req = FALSE) AND  (cancel = TRUE) AND  ( TRUE )) THEN
        cstate52 := 2; grant := FALSE;
    ELSIF ((req = TRUE) AND  (cancel = TRUE) AND  ( TRUE )) THEN
        cstate52 := 6; grant := FALSE;
    ELSIF ((req = TRUE) AND  (cancel = FALSE) AND  ( TRUE )) THEN
        cstate52 := 8; grant := TRUE;
    END_IF;
0:
    IF ((req = FALSE) AND  (cancel = FALSE) AND  ( TRUE )) THEN
        cstate52 := 25; grant := FALSE;
    ELSIF ((req = TRUE) AND  (cancel = FALSE) AND  ( TRUE )) THEN
        cstate52 := 4; grant := FALSE;
    ELSIF ((req = FALSE) AND  (cancel = TRUE) AND  ( TRUE )) THEN
        cstate52 := 20; grant := FALSE;
    ELSIF ((req = TRUE) AND  (cancel = TRUE) AND  ( TRUE )) THEN
        cstate52 := 16; grant := FALSE;
    END_IF;
1:
    IF ((req = FALSE) AND  (cancel = TRUE) AND  ( TRUE )) THEN
        cstate52 := 2; grant := FALSE;
    ELSIF ((req = FALSE) AND  (cancel = FALSE) AND  ( TRUE )) THEN
        cstate52 := 7; grant := FALSE;
    ELSIF ((req = TRUE) AND  (cancel = TRUE) AND  ( TRUE )) THEN
        cstate52 := 6; grant := FALSE;
    ELSIF ((req = TRUE) AND  (cancel = FALSE) AND  ( TRUE )) THEN
        cstate52 := 12; grant := FALSE;
    END_IF;
2:
    IF ((req = FALSE) AND  ( TRUE ) AND  (go = FALSE)) THEN
        cstate52 := 3; grant := FALSE;
    ELSIF ((req = TRUE) AND  ( TRUE ) AND  (go = FALSE)) THEN
        cstate52 := 21; grant := FALSE;
    ELSIF ((req = FALSE) AND  (cancel = FALSE) AND  (go = TRUE)) THEN
        cstate52 := 9; grant := FALSE;
    ELSIF ((req = FALSE) AND  (cancel = TRUE) AND  (go = TRUE)) THEN
        cstate52 := 2; grant := FALSE;
    ELSIF ((req = TRUE) AND  (cancel = FALSE) AND  (go = TRUE)) THEN
        cstate52 := 1; grant := FALSE;
    ELSIF ((req = TRUE) AND  (cancel = TRUE) AND  (go = TRUE)) THEN
        cstate52 := 6; grant := FALSE;
    END_IF;
3:
    IF ((req = TRUE) AND  (cancel = FALSE) AND  (go = TRUE)) THEN
        cstate52 := 4; grant := FALSE;
    ELSIF ((req = FALSE) AND  (cancel = TRUE) AND  (go = TRUE)) THEN
        cstate52 := 20; grant := FALSE;
    ELSIF ((req = TRUE) AND  (cancel = TRUE) AND  (go = TRUE)) THEN
        cstate52 := 16; grant := FALSE;
    ELSIF (( TRUE ) AND  ( TRUE ) AND  (go = FALSE)) THEN
        cstate52 := 22; grant := FALSE;
    ELSIF ((req = FALSE) AND  (cancel = FALSE) AND  (go = TRUE)) THEN
        cstate52 := 25; grant := FALSE;
    END_IF;
4:
    IF ((req = TRUE) AND  (cancel = FALSE) AND  ( TRUE )) THEN
        cstate52 := 12; grant := FALSE;
    ELSIF ((req = FALSE) AND  (cancel = FALSE) AND  ( TRUE )) THEN
        cstate52 := 7; grant := FALSE;
    ELSIF ((req = TRUE) AND  (cancel = TRUE) AND  ( TRUE )) THEN
        cstate52 := 6; grant := FALSE;
    ELSIF ((req = FALSE) AND  (cancel = TRUE) AND  ( TRUE )) THEN
        cstate52 := 2; grant := FALSE;
    END_IF;
5:
    IF ((req = TRUE) AND  (cancel = TRUE) AND  ( TRUE )) THEN
        cstate52 := 6; grant := FALSE;
    ELSIF ((req = FALSE) AND  (cancel = TRUE) AND  ( TRUE )) THEN
        cstate52 := 2; grant := FALSE;
    ELSIF ((req = FALSE) AND  (cancel = FALSE) AND  ( TRUE )) THEN
        cstate52 := 18; grant := TRUE;
    ELSIF ((req = TRUE) AND  (cancel = FALSE) AND  ( TRUE )) THEN
        cstate52 := 8; grant := TRUE;
    END_IF;
6:
    IF ((req = FALSE) AND  (cancel = TRUE) AND  (go = FALSE)) THEN
        cstate52 := 3; grant := FALSE;
    ELSIF ((req = TRUE) AND  (cancel = TRUE) AND  (go = TRUE)) THEN
        cstate52 := 6; grant := FALSE;
    ELSIF ((req = FALSE) AND  (cancel = FALSE) AND  (go = TRUE)) THEN
        cstate52 := 7; grant := FALSE;
    ELSIF ((req = TRUE) AND  (cancel = FALSE) AND  (go = FALSE)) THEN
        cstate52 := 10; grant := FALSE;
    ELSIF ((req = FALSE) AND  (cancel = TRUE) AND  (go = TRUE)) THEN
        cstate52 := 2; grant := FALSE;
    ELSIF ((req = TRUE) AND  (cancel = FALSE) AND  (go = TRUE)) THEN
        cstate52 := 12; grant := FALSE;
    ELSIF ((req = TRUE) AND  (cancel = TRUE) AND  (go = FALSE)) THEN
        cstate52 := 21; grant := FALSE;
    ELSIF ((req = FALSE) AND  (cancel = FALSE) AND  (go = FALSE)) THEN
        cstate52 := 27; grant := FALSE;
    END_IF;
7:
    IF ((req = FALSE) AND  (cancel = TRUE) AND  ( TRUE )) THEN
        cstate52 := 2; grant := FALSE;
    ELSIF ((req = TRUE) AND  (cancel = TRUE) AND  ( TRUE )) THEN
        cstate52 := 6; grant := FALSE;
    ELSIF ((req = TRUE) AND  (cancel = FALSE) AND  ( TRUE )) THEN
        cstate52 := 24; grant := FALSE;
    ELSIF ((req = FALSE) AND  (cancel = FALSE) AND  ( TRUE )) THEN
        cstate52 := 5; grant := FALSE;
    END_IF;
8:
    IF ((req = TRUE) AND  (cancel = TRUE) AND  ( TRUE )) THEN
        cstate52 := 6; grant := FALSE;
    ELSIF ((req = FALSE) AND  (cancel = FALSE) AND  ( TRUE )) THEN
        cstate52 := 7; grant := FALSE;
    ELSIF ((req = TRUE) AND  (cancel = FALSE) AND  ( TRUE )) THEN
        cstate52 := 12; grant := FALSE;
    ELSIF ((req = FALSE) AND  (cancel = TRUE) AND  ( TRUE )) THEN
        cstate52 := 2; grant := FALSE;
    END_IF;
9:
    IF ((req = FALSE) AND  (cancel = FALSE) AND  ( TRUE )) THEN
        cstate52 := 9; grant := FALSE;
    ELSIF ((req = TRUE) AND  (cancel = FALSE) AND  ( TRUE )) THEN
        cstate52 := 1; grant := FALSE;
    ELSIF ((req = TRUE) AND  (cancel = TRUE) AND  ( TRUE )) THEN
        cstate52 := 6; grant := FALSE;
    ELSIF ((req = FALSE) AND  (cancel = TRUE) AND  ( TRUE )) THEN
        cstate52 := 2; grant := FALSE;
    END_IF;
20:
    IF ((req = FALSE) AND  (cancel = TRUE) AND  (go = TRUE)) THEN
        cstate52 := 2; grant := FALSE;
    ELSIF ((req = TRUE) AND  ( TRUE ) AND  (go = FALSE)) THEN
        cstate52 := 21; grant := FALSE;
    ELSIF ((req = FALSE) AND  (cancel = FALSE) AND  (go = TRUE)) THEN
        cstate52 := 9; grant := FALSE;
    ELSIF ((req = FALSE) AND  ( TRUE ) AND  (go = FALSE)) THEN
        cstate52 := 3; grant := FALSE;
    ELSIF ((req = TRUE) AND  (cancel = FALSE) AND  (go = TRUE)) THEN
        cstate52 := 1; grant := FALSE;
    ELSIF ((req = TRUE) AND  (cancel = TRUE) AND  (go = TRUE)) THEN
        cstate52 := 6; grant := FALSE;
    END_IF;
21:
    IF ((req = TRUE) AND  (cancel = FALSE) AND  (go = TRUE)) THEN
        cstate52 := 14; grant := FALSE;
    ELSIF (( TRUE ) AND  ( TRUE ) AND  (go = FALSE)) THEN
        cstate52 := 22; grant := FALSE;
    ELSIF ((req = FALSE) AND  (cancel = TRUE) AND  (go = TRUE)) THEN
        cstate52 := 20; grant := FALSE;
    ELSIF ((req = FALSE) AND  (cancel = FALSE) AND  (go = TRUE)) THEN
        cstate52 := 23; grant := FALSE;
    ELSIF ((req = TRUE) AND  (cancel = TRUE) AND  (go = TRUE)) THEN
        cstate52 := 16; grant := FALSE;
    END_IF;
END_CASE;

END_FUNCTION_BLOCK
